(* IEC 61131-3 sources: TIA2AX/tests/V19/test_projects/expected/HW_2200330/ST80_PLC, 7 files *)

(* ---- HwIdentifiers.st ---- *)
TYPE
	HwIdentifiers : WORD
	(
		ST80_PLC_Profilschiene_0 :=	WORD#256,
		ST80_PLC :=	WORD#48,
		ST80_PLC_Card_reader_writer_1 :=	WORD#51,
		ST80_PLC_CPU_display_1 :=	WORD#54,
		ST80_PLC_OPC_UA_1 :=	WORD#117,
		ST80_PLC_DP_interface_1 :=	WORD#60,
		ST80_PLC_PROFINET_interface_1 :=	WORD#64,
		ST80_PLC_PROFINET_interface_1_Port_1 :=	WORD#65,
		ST80_PLC_PROFINET_interface_1_Port_2 :=	WORD#66,
		ST80_PLC_PROFINET_interface_2 :=	WORD#72,
		ST80_PLC_PROFINET_interface_2_Port_1 :=	WORD#73,
		ST80_Switch_SCALANCE_X_rack :=	WORD#412,
		ST80_Switch :=	WORD#413,
		ST80_Switch_ST80_Switch :=	WORD#414,
		ST80_Switch_SCALANCE_interface_1 :=	WORD#415,
		ST80_Switch_SCALANCE_interface_1_Port_1 :=	WORD#416,
		ST80_Switch_SCALANCE_interface_1_Port_2 :=	WORD#417,
		ST80_Switch_SCALANCE_interface_1_Port_3 :=	WORD#418,
		ST80_Switch_SCALANCE_interface_1_Port_4 :=	WORD#419,
		ST80_Switch_SCALANCE_interface_1_Port_5 :=	WORD#420,
		ST80_Switch_SCALANCE_interface_1_Port_6 :=	WORD#421,
		ST80_Switch_SCALANCE_interface_1_Port_7 :=	WORD#422,
		ST80_Switch_SCALANCE_interface_1_Port_8 :=	WORD#423,
		ST80_Switch_SCALANCE_interface_1_Port_9 :=	WORD#424,
		ST80_Switch_SCALANCE_interface_1_Port_10 :=	WORD#425,
		ST80_Switch_SCALANCE_interface_1_Port_11 :=	WORD#426,
		ST80_Switch_SCALANCE_interface_1_Port_12 :=	WORD#427,
		ST80_Switch_SCALANCE_interface_1_Port_13 :=	WORD#428,
		ST80_Switch_SCALANCE_interface_1_Port_14 :=	WORD#429,
		ST80_Switch_SCALANCE_interface_1_Port_15 :=	WORD#430,
		ST80_Switch_SCALANCE_interface_1_Port_16 :=	WORD#431,
		ST80_1_DM260_EB_Box_Rack :=	WORD#270,
		ST80_1_DM260_EB_Box :=	WORD#258,
		ST80_1_DM260_EB_Box_Interface :=	WORD#259,
		ST80_1_DM260_EB_Box_Interface_Port_1 :=	WORD#260,
		ST80_1_DM260_EB_Box_DataMan_260 :=	WORD#261,
		ST80_1_DM260_EB_Box_Acquisition_Control_1 :=	WORD#262,
		ST80_1_DM260_EB_Box_Acquisition_Status_1 :=	WORD#263,
		ST80_1_DM260_EB_Box_Results_Control_1 :=	WORD#264,
		ST80_1_DM260_EB_Box_Results_Status_1 :=	WORD#265,
		ST80_1_DM260_EB_Box_Soft_Event_Control_1 :=	WORD#266,
		ST80_1_DM260_EB_Box_User_Data_64_bytes_1 :=	WORD#267,
		ST80_1_DM260_EB_Box_Result_Data_64_bytes_1 :=	WORD#268,
		ST80_HMI_ConnectionBox_2_Connection_Box :=	WORD#272,
		ST80_HMI_ConnectionBox_2 :=	WORD#273,
		ST80_HMI_ConnectionBox_2_ST80_HMI_ConnectionBox_2 :=	WORD#274,
		ST80_HMI_ConnectionBox_2_SCALANCE_interface_1 :=	WORD#275,
		ST80_HMI_ConnectionBox_2_SCALANCE_interface_1_Port_1 :=	WORD#276,
		ST80_HMI_ConnectionBox_2_SCALANCE_interface_1_Port_2 :=	WORD#277,
		ST80_HMI_ConnectionBox_2_SCALANCE_interface_1_Port_3 :=	WORD#278,
		ST80_1_CMMT_1GF1_PN_IO_Interface :=	WORD#282,
		ST80_1_CMMT_1GF1_PN_IO_Interface_Port_1 :=	WORD#283,
		ST80_1_CMMT_1GF1_PN_IO_Interface_Port_2 :=	WORD#284,
		ST80_1_CMMT_1GF1_CMMT_AS_V1 :=	WORD#285,
		ST80_1_CMMT_1GF1_DO_SERVO_1_Module_Access_Point :=	WORD#287,
		ST80_1_CMMT_1GF1_DO_SERVO_1_Siemens_telegram_111_PZD_12_12 :=	WORD#288,
		ST80_1_CMMT_1GF1_Siemens_telegram_111_PZD_12_12 :=	WORD#288,
		ST80_1_CMMT_1GF2_PN_IO_Interface :=	WORD#292,
		ST80_1_CMMT_1GF2_PN_IO_Interface_Port_1 :=	WORD#293,
		ST80_1_CMMT_1GF2_PN_IO_Interface_Port_2 :=	WORD#294,
		ST80_1_CMMT_1GF2_CMMT_AS_V1 :=	WORD#295,
		ST80_1_CMMT_1GF2_DO_SERVO_1_Module_Access_Point :=	WORD#297,
		ST80_1_CMMT_1GF2_DO_SERVO_1_Siemens_telegram_111_PZD_12_12 :=	WORD#298,
		ST80_1_CMMT_1GF2_Siemens_telegram_111_PZD_12_12 :=	WORD#298,
		ST80_1_DM260_PB_Box_Rack :=	WORD#300,
		ST80_1_DM260_PB_Box :=	WORD#301,
		ST80_1_DM260_PB_Box_Interface :=	WORD#302,
		ST80_1_DM260_PB_Box_Interface_Port_1 :=	WORD#303,
		ST80_1_DM260_PB_Box_DataMan_260 :=	WORD#304,
		ST80_1_DM260_PB_Box_Acquisition_Control_1 :=	WORD#305,
		ST80_1_DM260_PB_Box_Acquisition_Status_1 :=	WORD#306,
		ST80_1_DM260_PB_Box_Results_Control_1 :=	WORD#307,
		ST80_1_DM260_PB_Box_Results_Status_1 :=	WORD#308,
		ST80_1_DM260_PB_Box_Soft_Event_Control_1 :=	WORD#309,
		ST80_1_DM260_PB_Box_User_Data_64_bytes_1 :=	WORD#310,
		ST80_1_DM260_PB_Box_Result_Data_64_bytes_1 :=	WORD#311,
		ST80_ET200SP_2_Rack_0 :=	WORD#313,
		ST80_ET200SP_2 :=	WORD#314,
		ST80_ET200SP_2_ST80_ET200SP_2 :=	WORD#315,
		ST80_ET200SP_2_PROFINET_interface :=	WORD#316,
		ST80_ET200SP_2_PROFINET_interface_Port_1 :=	WORD#318,
		ST80_ET200SP_2_PROFINET_interface_Port_2 :=	WORD#317,
		ST80_ET200SP_2_BA_2xRJ45 :=	WORD#318,
		ST80_ET200SP_2_BU_Cover_15_mm_1 :=	WORD#319,
		ST80_ET200SP_2_11M1 :=	WORD#320,
		ST80_ET200SP_2_11M2 :=	WORD#321,
		ST80_ET200SP_2_11M3 :=	WORD#322,
		ST80_ET200SP_2_11M4 :=	WORD#323,
		ST80_ET200SP_2_12M1 :=	WORD#324,
		ST80_ET200SP_2_12M2 :=	WORD#325,
		ST80_ET200SP_2_12M3 :=	WORD#326,
		ST80_ET200SP_2_12M4 :=	WORD#327,
		ST80_ET200SP_2_13M1 :=	WORD#328,
		ST80_ET200SP_2_13M2 :=	WORD#329,
		ST80_ET200SP_2_13M3 :=	WORD#330,
		ST80_ET200SP_2_13M4 :=	WORD#331,
		ST80_ET200SP_2_Servermodul_1 :=	WORD#332,
		ST80_1_TZ535_PN_Rack :=	WORD#334,
		ST80_1_TZ535_PN :=	WORD#335,
		ST80_1_TZ535_PN_Interface :=	WORD#336,
		ST80_1_TZ535_PN_Interface_Port_1 :=	WORD#337,
		ST80_1_TZ535_PN_Interface_Port_2 :=	WORD#338,
		ST80_1_TZ535_PN_2D_TZ535_PN_PROFINET_IO :=	WORD#339,
		ST80_1_TZ535_PN_In_Out_32_byte_1 :=	WORD#340,
		ST80_1_DM260_Housing_Rack :=	WORD#342,
		ST80_1_DM260_Housing :=	WORD#343,
		ST80_1_DM260_Housing_Interface :=	WORD#344,
		ST80_1_DM260_Housing_Interface_Port_1 :=	WORD#345,
		ST80_1_DM260_Housing_DataMan_260 :=	WORD#346,
		ST80_1_DM260_Housing_Acquisition_Control_1 :=	WORD#347,
		ST80_1_DM260_Housing_Acquisition_Status_1 :=	WORD#348,
		ST80_1_DM260_Housing_Results_Control_1 :=	WORD#349,
		ST80_1_DM260_Housing_Results_Status_1 :=	WORD#350,
		ST80_1_DM260_Housing_Soft_Event_Control_1 :=	WORD#351,
		ST80_1_DM260_Housing_User_Data_64_bytes_1 :=	WORD#352,
		ST80_1_DM260_Housing_Result_Data_64_bytes_1 :=	WORD#353,
		ST80_1_CMMT_3GF1_PN_IO_Interface :=	WORD#357,
		ST80_1_CMMT_3GF1_PN_IO_Interface_Port_1 :=	WORD#358,
		ST80_1_CMMT_3GF1_PN_IO_Interface_Port_2 :=	WORD#359,
		ST80_1_CMMT_3GF1_CMMT_AS_V1 :=	WORD#360,
		ST80_1_CMMT_3GF1_DO_SERVO_1_Module_Access_Point :=	WORD#362,
		ST80_1_CMMT_3GF1_DO_SERVO_1_Siemens_telegram_111_PZD_12_12 :=	WORD#363,
		ST80_1_CMMT_3GF1_Siemens_telegram_111_PZD_12_12 :=	WORD#363,
		ST80_CPX_PN_IO_Interface :=	WORD#367,
		ST80_CPX_PN_IO_Interface_Port_1 :=	WORD#368,
		ST80_CPX_PN_IO_Interface_Port_2 :=	WORD#369,
		ST80_CPX_CPX :=	WORD#370,
		ST80_CPX_MPA1S_VMPA1_FB_EMS_8_8DO_1 :=	WORD#371,
		ST80_CPX_MPA1S_VMPA1_FB_EMS_8_8DO_2 :=	WORD#372,
		ST80_CPX_MPA2S_VMPA2_FB_EMS_4_4DO_1 :=	WORD#373,
		ST80_CPX_MPA1S_VMPA1_FB_EMS_8_8DO_3 :=	WORD#374,
		ST80_CPX_MPA2S_VMPA2_FB_EMS_4_4DO_2 :=	WORD#375,
		ST80_CPX_MPA1S_VMPA1_FB_EMS_8_8DO_4 :=	WORD#376,
		ST80_CPX_MPA1S_VMPA1_FB_EMS_8_8DO_5 :=	WORD#377,
		ST80_CPX_MPA1G_VMPA1_FB_EMG_8_8DO_1 :=	WORD#378,
		ST80_CPX_MPA1G_VMPA1_FB_EMG_8_8DO_2 :=	WORD#379,
		ST80_CPX_MPA2G_VMPA2_FB_EMG_4_4DO_1 :=	WORD#380,
		ST80_CPX_MPA1G_VMPA1_FB_EMG_8_8DO_3 :=	WORD#381,
		ST80_CPX_MPA1G_VMPA1_FB_EMG_8_8DO_4 :=	WORD#382,
		ST80_CPX_MPA1G_VMPA1_FB_EMG_8_8DO_5 :=	WORD#383,
		ST80_CPX_MPA1G_VMPA1_FB_EMG_8_8DO_6 :=	WORD#384,
		ST80_ET200SP_Rack_0 :=	WORD#386,
		ST80_ET200SP :=	WORD#387,
		ST80_ET200SP_ST80_ET200SP :=	WORD#388,
		ST80_ET200SP_PROFINET_interface :=	WORD#389,
		ST80_ET200SP_PROFINET_interface_Port_1 :=	WORD#391,
		ST80_ET200SP_PROFINET_interface_Port_2 :=	WORD#390,
		ST80_ET200SP_BA_2xRJ45 :=	WORD#391,
		ST80_ET200SP_CM_4xIO_Link_1 :=	WORD#392,
		ST80_ET200SP_CM_4xIO_Link_2 :=	WORD#393,
		ST80_ET200SP_CM_4xIO_Link_3 :=	WORD#394,
		ST80_ET200SP_DI_16x24VDC_ST_1 :=	WORD#395,
		ST80_ET200SP_DI_16x24VDC_ST_2 :=	WORD#396,
		ST80_ET200SP_DI_16x24VDC_ST_3 :=	WORD#397,
		ST80_ET200SP_DI_16x24VDC_ST_4 :=	WORD#398,
		ST80_ET200SP_DQ_16x24VDC_0_5A_ST_1 :=	WORD#399,
		ST80_ET200SP_DQ_16x24VDC_0_5A_ST_2 :=	WORD#400,
		ST80_ET200SP_DQ_16x24VDC_0_5A_ST_3 :=	WORD#401,
		ST80_ET200SP_Servermodul_1 :=	WORD#402,
		ST80_HMI_ConnectionBox_Connection_Box :=	WORD#404,
		ST80_HMI_ConnectionBox :=	WORD#405,
		ST80_HMI_ConnectionBox_ST80_HMI_ConnectionBox :=	WORD#406,
		ST80_HMI_ConnectionBox_SCALANCE_interface_1 :=	WORD#407,
		ST80_HMI_ConnectionBox_SCALANCE_interface_1_Port_1 :=	WORD#408,
		ST80_HMI_ConnectionBox_SCALANCE_interface_1_Port_2 :=	WORD#409,
		ST80_HMI_ConnectionBox_SCALANCE_interface_1_Port_3 :=	WORD#410,
		NONE:= WORD#0
	);
END_TYPE

(* ---- HwInputs.st ---- *)
TYPE
	HwInputs : STRUCT
		ST80_1_DM260_EB_Box_Acquisition_Status_1 AT %B1205 : ARRAY[0..2] OF BYTE;
		ST80_1_DM260_EB_Box_Results_Status_1 AT %B1208 : BYTE;
		ST80_1_DM260_EB_Box_Soft_Event_Control_1 AT %B1209 : BYTE;
		ST80_1_DM260_EB_Box_Result_Data_64_bytes_1 AT %B1382 : ARRAY[0..71] OF BYTE;
		ST80_1_CMMT_1GF1_DO_SERVO_1_Siemens_telegram_111_PZD_12_12 AT %B1700 : ARRAY[0..23] OF BYTE;
		ST80_1_CMMT_1GF2_DO_SERVO_1_Siemens_telegram_111_PZD_12_12 AT %B1600 : ARRAY[0..23] OF BYTE;
		ST80_1_DM260_PB_Box_Acquisition_Status_1 AT %B1200 : ARRAY[0..2] OF BYTE;
		ST80_1_DM260_PB_Box_Results_Status_1 AT %B1203 : BYTE;
		ST80_1_DM260_PB_Box_Soft_Event_Control_1 AT %B1204 : BYTE;
		ST80_1_DM260_PB_Box_Result_Data_64_bytes_1 AT %B1210 : ARRAY[0..71] OF BYTE;
		ST80_ET200SP_2_11M1 AT %B600 : DWORD;
		ST80_ET200SP_2_11M2 AT %B604 : DWORD;
		ST80_ET200SP_2_11M3 AT %B608 : DWORD;
		ST80_ET200SP_2_11M4 AT %B612 : DWORD;
		ST80_ET200SP_2_12M1 AT %B616 : DWORD;
		ST80_ET200SP_2_12M2 AT %B620 : DWORD;
		ST80_ET200SP_2_12M3 AT %B624 : DWORD;
		ST80_ET200SP_2_12M4 AT %B628 : DWORD;
		ST80_ET200SP_2_13M1 AT %B632 : DWORD;
		ST80_ET200SP_2_13M2 AT %B636 : DWORD;
		ST80_ET200SP_2_13M3 AT %B640 : DWORD;
		ST80_ET200SP_2_13M4 AT %B644 : DWORD;
		ST80_1_TZ535_PN_In_Out_32_byte_1 AT %B1800 : ARRAY[0..31] OF BYTE;
		ST80_1_DM260_Housing_Acquisition_Status_1 AT %B1000 : ARRAY[0..2] OF BYTE;
		ST80_1_DM260_Housing_Results_Status_1 AT %B1003 : BYTE;
		ST80_1_DM260_Housing_Soft_Event_Control_1 AT %B1004 : BYTE;
		ST80_1_DM260_Housing_Result_Data_64_bytes_1 AT %B1010 : ARRAY[0..71] OF BYTE;
		ST80_1_CMMT_3GF1_DO_SERVO_1_Siemens_telegram_111_PZD_12_12 AT %B1500 : ARRAY[0..23] OF BYTE;
		ST80_ET200SP_CM_4xIO_Link_1 AT %B100 : ARRAY[0..31] OF BYTE;
		ST80_ET200SP_CM_4xIO_Link_2 AT %B132 : ARRAY[0..31] OF BYTE;
		ST80_ET200SP_CM_4xIO_Link_3 AT %B164 : ARRAY[0..31] OF BYTE;
		ST80_ET200SP_DI_16x24VDC_ST_1 AT %B0 : WORD;
		ST80_ET200SP_DI_16x24VDC_ST_2 AT %B2 : WORD;
		ST80_ET200SP_DI_16x24VDC_ST_3 AT %B4 : WORD;
		ST80_ET200SP_DI_16x24VDC_ST_4 AT %B6 : WORD;
	END_STRUCT;
END_TYPE

(* ---- HwOutputs.st ---- *)
TYPE
	HwOutputs : STRUCT
		ST80_1_DM260_EB_Box_Acquisition_Control_1 AT %B1201 : BYTE;
		ST80_1_DM260_EB_Box_Results_Control_1 AT %B1205 : BYTE;
		ST80_1_DM260_EB_Box_Soft_Event_Control_1 AT %B1206 : BYTE;
		ST80_1_DM260_EB_Box_User_Data_64_bytes_1 AT %B1378 : ARRAY[0..67] OF BYTE;
		ST80_1_CMMT_1GF1_DO_SERVO_1_Siemens_telegram_111_PZD_12_12 AT %B1700 : ARRAY[0..23] OF BYTE;
		ST80_1_CMMT_1GF2_DO_SERVO_1_Siemens_telegram_111_PZD_12_12 AT %B1600 : ARRAY[0..23] OF BYTE;
		ST80_1_DM260_PB_Box_Acquisition_Control_1 AT %B1200 : BYTE;
		ST80_1_DM260_PB_Box_Results_Control_1 AT %B1203 : BYTE;
		ST80_1_DM260_PB_Box_Soft_Event_Control_1 AT %B1204 : BYTE;
		ST80_1_DM260_PB_Box_User_Data_64_bytes_1 AT %B1210 : ARRAY[0..67] OF BYTE;
		ST80_ET200SP_2_11M1 AT %B600 : WORD;
		ST80_ET200SP_2_11M2 AT %B604 : WORD;
		ST80_ET200SP_2_11M3 AT %B608 : WORD;
		ST80_ET200SP_2_11M4 AT %B612 : WORD;
		ST80_ET200SP_2_12M1 AT %B616 : WORD;
		ST80_ET200SP_2_12M2 AT %B620 : WORD;
		ST80_ET200SP_2_12M3 AT %B624 : WORD;
		ST80_ET200SP_2_12M4 AT %B628 : WORD;
		ST80_ET200SP_2_13M1 AT %B632 : WORD;
		ST80_ET200SP_2_13M2 AT %B636 : WORD;
		ST80_ET200SP_2_13M3 AT %B640 : WORD;
		ST80_ET200SP_2_13M4 AT %B644 : WORD;
		ST80_1_TZ535_PN_In_Out_32_byte_1 AT %B1800 : ARRAY[0..31] OF BYTE;
		ST80_1_DM260_Housing_Acquisition_Control_1 AT %B1000 : BYTE;
		ST80_1_DM260_Housing_Results_Control_1 AT %B1003 : BYTE;
		ST80_1_DM260_Housing_Soft_Event_Control_1 AT %B1004 : BYTE;
		ST80_1_DM260_Housing_User_Data_64_bytes_1 AT %B1010 : ARRAY[0..67] OF BYTE;
		ST80_1_CMMT_3GF1_DO_SERVO_1_Siemens_telegram_111_PZD_12_12 AT %B1500 : ARRAY[0..23] OF BYTE;
		ST80_CPX_MPA1S_VMPA1_FB_EMS_8_8DO_1 AT %B200 : BYTE;
		ST80_CPX_MPA1S_VMPA1_FB_EMS_8_8DO_2 AT %B201 : BYTE;
		ST80_CPX_MPA2S_VMPA2_FB_EMS_4_4DO_1 AT %B202 : BYTE;
		ST80_CPX_MPA1S_VMPA1_FB_EMS_8_8DO_3 AT %B203 : BYTE;
		ST80_CPX_MPA2S_VMPA2_FB_EMS_4_4DO_2 AT %B204 : BYTE;
		ST80_CPX_MPA1S_VMPA1_FB_EMS_8_8DO_4 AT %B205 : BYTE;
		ST80_CPX_MPA1S_VMPA1_FB_EMS_8_8DO_5 AT %B206 : BYTE;
		ST80_CPX_MPA1G_VMPA1_FB_EMG_8_8DO_1 AT %B207 : BYTE;
		ST80_CPX_MPA1G_VMPA1_FB_EMG_8_8DO_2 AT %B208 : BYTE;
		ST80_CPX_MPA2G_VMPA2_FB_EMG_4_4DO_1 AT %B209 : BYTE;
		ST80_CPX_MPA1G_VMPA1_FB_EMG_8_8DO_3 AT %B210 : BYTE;
		ST80_CPX_MPA1G_VMPA1_FB_EMG_8_8DO_4 AT %B211 : BYTE;
		ST80_CPX_MPA1G_VMPA1_FB_EMG_8_8DO_5 AT %B212 : BYTE;
		ST80_CPX_MPA1G_VMPA1_FB_EMG_8_8DO_6 AT %B213 : BYTE;
		ST80_ET200SP_CM_4xIO_Link_1 AT %B100 : ARRAY[0..31] OF BYTE;
		ST80_ET200SP_CM_4xIO_Link_2 AT %B132 : ARRAY[0..31] OF BYTE;
		ST80_ET200SP_CM_4xIO_Link_3 AT %B164 : ARRAY[0..31] OF BYTE;
		ST80_ET200SP_DQ_16x24VDC_0_5A_ST_1 AT %B0 : WORD;
		ST80_ET200SP_DQ_16x24VDC_0_5A_ST_2 AT %B2 : WORD;
		ST80_ET200SP_DQ_16x24VDC_0_5A_ST_3 AT %B4 : WORD;
	END_STRUCT;
END_TYPE

(* ---- PlcInputs.st ---- *)
TYPE
	PlcInputs : STRUCT
		ST80_1_DM260_EB_Box_Acquisition_Status_1 : ARRAY[0..2] OF BYTE;
		ST80_1_DM260_EB_Box_Results_Status_1 : BYTE;
		ST80_1_DM260_EB_Box_Soft_Event_Control_1 : BYTE;
		ST80_1_DM260_EB_Box_Result_Data_64_bytes_1 : ARRAY[0..71] OF BYTE;
		ST80_1_CMMT_1GF1_DO_SERVO_1_Siemens_telegram_111_PZD_12_12 : ARRAY[0..23] OF BYTE;
		ST80_1_CMMT_1GF2_DO_SERVO_1_Siemens_telegram_111_PZD_12_12 : ARRAY[0..23] OF BYTE;
		ST80_1_DM260_PB_Box_Acquisition_Status_1 : ARRAY[0..2] OF BYTE;
		ST80_1_DM260_PB_Box_Results_Status_1 : BYTE;
		ST80_1_DM260_PB_Box_Soft_Event_Control_1 : BYTE;
		ST80_1_DM260_PB_Box_Result_Data_64_bytes_1 : ARRAY[0..71] OF BYTE;
		ST80_ET200SP_2_11M1 : DWORD;
		ST80_ET200SP_2_11M2 : DWORD;
		ST80_ET200SP_2_11M3 : DWORD;
		ST80_ET200SP_2_11M4 : DWORD;
		ST80_ET200SP_2_12M1 : DWORD;
		ST80_ET200SP_2_12M2 : DWORD;
		ST80_ET200SP_2_12M3 : DWORD;
		ST80_ET200SP_2_12M4 : DWORD;
		ST80_ET200SP_2_13M1 : DWORD;
		ST80_ET200SP_2_13M2 : DWORD;
		ST80_ET200SP_2_13M3 : DWORD;
		ST80_ET200SP_2_13M4 : DWORD;
		ST80_1_TZ535_PN_In_Out_32_byte_1 : ARRAY[0..31] OF BYTE;
		ST80_1_DM260_Housing_Acquisition_Status_1 : ARRAY[0..2] OF BYTE;
		ST80_1_DM260_Housing_Results_Status_1 : BYTE;
		ST80_1_DM260_Housing_Soft_Event_Control_1 : BYTE;
		ST80_1_DM260_Housing_Result_Data_64_bytes_1 : ARRAY[0..71] OF BYTE;
		ST80_1_CMMT_3GF1_DO_SERVO_1_Siemens_telegram_111_PZD_12_12 : ARRAY[0..23] OF BYTE;
		ST80_ET200SP_CM_4xIO_Link_1 : ARRAY[0..31] OF BYTE;
		ST80_ET200SP_CM_4xIO_Link_2 : ARRAY[0..31] OF BYTE;
		ST80_ET200SP_CM_4xIO_Link_3 : ARRAY[0..31] OF BYTE;
		ST80_ET200SP_DI_16x24VDC_ST_1 : WORD;
		ST80_ET200SP_DI_16x24VDC_ST_2 : WORD;
		ST80_ET200SP_DI_16x24VDC_ST_3 : WORD;
		ST80_ET200SP_DI_16x24VDC_ST_4 : WORD;
	END_STRUCT;
END_TYPE

(* ---- PlcOutputs.st ---- *)
TYPE
	PlcOutputs : STRUCT
		ST80_1_DM260_EB_Box_Acquisition_Control_1 : BYTE;
		ST80_1_DM260_EB_Box_Results_Control_1 : BYTE;
		ST80_1_DM260_EB_Box_Soft_Event_Control_1 : BYTE;
		ST80_1_DM260_EB_Box_User_Data_64_bytes_1 : ARRAY[0..67] OF BYTE;
		ST80_1_CMMT_1GF1_DO_SERVO_1_Siemens_telegram_111_PZD_12_12 : ARRAY[0..23] OF BYTE;
		ST80_1_CMMT_1GF2_DO_SERVO_1_Siemens_telegram_111_PZD_12_12 : ARRAY[0..23] OF BYTE;
		ST80_1_DM260_PB_Box_Acquisition_Control_1 : BYTE;
		ST80_1_DM260_PB_Box_Results_Control_1 : BYTE;
		ST80_1_DM260_PB_Box_Soft_Event_Control_1 : BYTE;
		ST80_1_DM260_PB_Box_User_Data_64_bytes_1 : ARRAY[0..67] OF BYTE;
		ST80_ET200SP_2_11M1 : WORD;
		ST80_ET200SP_2_11M2 : WORD;
		ST80_ET200SP_2_11M3 : WORD;
		ST80_ET200SP_2_11M4 : WORD;
		ST80_ET200SP_2_12M1 : WORD;
		ST80_ET200SP_2_12M2 : WORD;
		ST80_ET200SP_2_12M3 : WORD;
		ST80_ET200SP_2_12M4 : WORD;
		ST80_ET200SP_2_13M1 : WORD;
		ST80_ET200SP_2_13M2 : WORD;
		ST80_ET200SP_2_13M3 : WORD;
		ST80_ET200SP_2_13M4 : WORD;
		ST80_1_TZ535_PN_In_Out_32_byte_1 : ARRAY[0..31] OF BYTE;
		ST80_1_DM260_Housing_Acquisition_Control_1 : BYTE;
		ST80_1_DM260_Housing_Results_Control_1 : BYTE;
		ST80_1_DM260_Housing_Soft_Event_Control_1 : BYTE;
		ST80_1_DM260_Housing_User_Data_64_bytes_1 : ARRAY[0..67] OF BYTE;
		ST80_1_CMMT_3GF1_DO_SERVO_1_Siemens_telegram_111_PZD_12_12 : ARRAY[0..23] OF BYTE;
		ST80_CPX_MPA1S_VMPA1_FB_EMS_8_8DO_1 : BYTE;
		ST80_CPX_MPA1S_VMPA1_FB_EMS_8_8DO_2 : BYTE;
		ST80_CPX_MPA2S_VMPA2_FB_EMS_4_4DO_1 : BYTE;
		ST80_CPX_MPA1S_VMPA1_FB_EMS_8_8DO_3 : BYTE;
		ST80_CPX_MPA2S_VMPA2_FB_EMS_4_4DO_2 : BYTE;
		ST80_CPX_MPA1S_VMPA1_FB_EMS_8_8DO_4 : BYTE;
		ST80_CPX_MPA1S_VMPA1_FB_EMS_8_8DO_5 : BYTE;
		ST80_CPX_MPA1G_VMPA1_FB_EMG_8_8DO_1 : BYTE;
		ST80_CPX_MPA1G_VMPA1_FB_EMG_8_8DO_2 : BYTE;
		ST80_CPX_MPA2G_VMPA2_FB_EMG_4_4DO_1 : BYTE;
		ST80_CPX_MPA1G_VMPA1_FB_EMG_8_8DO_3 : BYTE;
		ST80_CPX_MPA1G_VMPA1_FB_EMG_8_8DO_4 : BYTE;
		ST80_CPX_MPA1G_VMPA1_FB_EMG_8_8DO_5 : BYTE;
		ST80_CPX_MPA1G_VMPA1_FB_EMG_8_8DO_6 : BYTE;
		ST80_ET200SP_CM_4xIO_Link_1 : ARRAY[0..31] OF BYTE;
		ST80_ET200SP_CM_4xIO_Link_2 : ARRAY[0..31] OF BYTE;
		ST80_ET200SP_CM_4xIO_Link_3 : ARRAY[0..31] OF BYTE;
		ST80_ET200SP_DQ_16x24VDC_0_5A_ST_1 : WORD;
		ST80_ET200SP_DQ_16x24VDC_0_5A_ST_2 : WORD;
		ST80_ET200SP_DQ_16x24VDC_0_5A_ST_3 : WORD;
	END_STRUCT;
END_TYPE

(* ---- CopyInputs.st ---- *)
FUNCTION CopyInputs
	VAR_EXTERNAL
		HwInputs : HwInputs;
		PlcInputs : PlcInputs;
	END_VAR
	PlcInputs.ST80_1_DM260_EB_Box_Acquisition_Status_1[0] := HwInputs.ST80_1_DM260_EB_Box_Acquisition_Status_1[0];
	PlcInputs.ST80_1_DM260_EB_Box_Acquisition_Status_1[1] := HwInputs.ST80_1_DM260_EB_Box_Acquisition_Status_1[1];
	PlcInputs.ST80_1_DM260_EB_Box_Acquisition_Status_1[2] := HwInputs.ST80_1_DM260_EB_Box_Acquisition_Status_1[2];
	PlcInputs.ST80_1_DM260_EB_Box_Results_Status_1 := HwInputs.ST80_1_DM260_EB_Box_Results_Status_1;
	PlcInputs.ST80_1_DM260_EB_Box_Soft_Event_Control_1 := HwInputs.ST80_1_DM260_EB_Box_Soft_Event_Control_1;
	PlcInputs.ST80_1_DM260_EB_Box_Result_Data_64_bytes_1[0] := HwInputs.ST80_1_DM260_EB_Box_Result_Data_64_bytes_1[0];
	PlcInputs.ST80_1_DM260_EB_Box_Result_Data_64_bytes_1[1] := HwInputs.ST80_1_DM260_EB_Box_Result_Data_64_bytes_1[1];
	PlcInputs.ST80_1_DM260_EB_Box_Result_Data_64_bytes_1[2] := HwInputs.ST80_1_DM260_EB_Box_Result_Data_64_bytes_1[2];
	PlcInputs.ST80_1_DM260_EB_Box_Result_Data_64_bytes_1[3] := HwInputs.ST80_1_DM260_EB_Box_Result_Data_64_bytes_1[3];
	PlcInputs.ST80_1_DM260_EB_Box_Result_Data_64_bytes_1[4] := HwInputs.ST80_1_DM260_EB_Box_Result_Data_64_bytes_1[4];
	PlcInputs.ST80_1_DM260_EB_Box_Result_Data_64_bytes_1[5] := HwInputs.ST80_1_DM260_EB_Box_Result_Data_64_bytes_1[5];
	PlcInputs.ST80_1_DM260_EB_Box_Result_Data_64_bytes_1[6] := HwInputs.ST80_1_DM260_EB_Box_Result_Data_64_bytes_1[6];
	PlcInputs.ST80_1_DM260_EB_Box_Result_Data_64_bytes_1[7] := HwInputs.ST80_1_DM260_EB_Box_Result_Data_64_bytes_1[7];
	PlcInputs.ST80_1_DM260_EB_Box_Result_Data_64_bytes_1[8] := HwInputs.ST80_1_DM260_EB_Box_Result_Data_64_bytes_1[8];
	PlcInputs.ST80_1_DM260_EB_Box_Result_Data_64_bytes_1[9] := HwInputs.ST80_1_DM260_EB_Box_Result_Data_64_bytes_1[9];
	PlcInputs.ST80_1_DM260_EB_Box_Result_Data_64_bytes_1[10] := HwInputs.ST80_1_DM260_EB_Box_Result_Data_64_bytes_1[10];
	PlcInputs.ST80_1_DM260_EB_Box_Result_Data_64_bytes_1[11] := HwInputs.ST80_1_DM260_EB_Box_Result_Data_64_bytes_1[11];
	PlcInputs.ST80_1_DM260_EB_Box_Result_Data_64_bytes_1[12] := HwInputs.ST80_1_DM260_EB_Box_Result_Data_64_bytes_1[12];
	PlcInputs.ST80_1_DM260_EB_Box_Result_Data_64_bytes_1[13] := HwInputs.ST80_1_DM260_EB_Box_Result_Data_64_bytes_1[13];
	PlcInputs.ST80_1_DM260_EB_Box_Result_Data_64_bytes_1[14] := HwInputs.ST80_1_DM260_EB_Box_Result_Data_64_bytes_1[14];
	PlcInputs.ST80_1_DM260_EB_Box_Result_Data_64_bytes_1[15] := HwInputs.ST80_1_DM260_EB_Box_Result_Data_64_bytes_1[15];
	PlcInputs.ST80_1_DM260_EB_Box_Result_Data_64_bytes_1[16] := HwInputs.ST80_1_DM260_EB_Box_Result_Data_64_bytes_1[16];
	PlcInputs.ST80_1_DM260_EB_Box_Result_Data_64_bytes_1[17] := HwInputs.ST80_1_DM260_EB_Box_Result_Data_64_bytes_1[17];
	PlcInputs.ST80_1_DM260_EB_Box_Result_Data_64_bytes_1[18] := HwInputs.ST80_1_DM260_EB_Box_Result_Data_64_bytes_1[18];
	PlcInputs.ST80_1_DM260_EB_Box_Result_Data_64_bytes_1[19] := HwInputs.ST80_1_DM260_EB_Box_Result_Data_64_bytes_1[19];
	PlcInputs.ST80_1_DM260_EB_Box_Result_Data_64_bytes_1[20] := HwInputs.ST80_1_DM260_EB_Box_Result_Data_64_bytes_1[20];
	PlcInputs.ST80_1_DM260_EB_Box_Result_Data_64_bytes_1[21] := HwInputs.ST80_1_DM260_EB_Box_Result_Data_64_bytes_1[21];
	PlcInputs.ST80_1_DM260_EB_Box_Result_Data_64_bytes_1[22] := HwInputs.ST80_1_DM260_EB_Box_Result_Data_64_bytes_1[22];
	PlcInputs.ST80_1_DM260_EB_Box_Result_Data_64_bytes_1[23] := HwInputs.ST80_1_DM260_EB_Box_Result_Data_64_bytes_1[23];
	PlcInputs.ST80_1_DM260_EB_Box_Result_Data_64_bytes_1[24] := HwInputs.ST80_1_DM260_EB_Box_Result_Data_64_bytes_1[24];
	PlcInputs.ST80_1_DM260_EB_Box_Result_Data_64_bytes_1[25] := HwInputs.ST80_1_DM260_EB_Box_Result_Data_64_bytes_1[25];
	PlcInputs.ST80_1_DM260_EB_Box_Result_Data_64_bytes_1[26] := HwInputs.ST80_1_DM260_EB_Box_Result_Data_64_bytes_1[26];
	PlcInputs.ST80_1_DM260_EB_Box_Result_Data_64_bytes_1[27] := HwInputs.ST80_1_DM260_EB_Box_Result_Data_64_bytes_1[27];
	PlcInputs.ST80_1_DM260_EB_Box_Result_Data_64_bytes_1[28] := HwInputs.ST80_1_DM260_EB_Box_Result_Data_64_bytes_1[28];
	PlcInputs.ST80_1_DM260_EB_Box_Result_Data_64_bytes_1[29] := HwInputs.ST80_1_DM260_EB_Box_Result_Data_64_bytes_1[29];
	PlcInputs.ST80_1_DM260_EB_Box_Result_Data_64_bytes_1[30] := HwInputs.ST80_1_DM260_EB_Box_Result_Data_64_bytes_1[30];
	PlcInputs.ST80_1_DM260_EB_Box_Result_Data_64_bytes_1[31] := HwInputs.ST80_1_DM260_EB_Box_Result_Data_64_bytes_1[31];
	PlcInputs.ST80_1_DM260_EB_Box_Result_Data_64_bytes_1[32] := HwInputs.ST80_1_DM260_EB_Box_Result_Data_64_bytes_1[32];
	PlcInputs.ST80_1_DM260_EB_Box_Result_Data_64_bytes_1[33] := HwInputs.ST80_1_DM260_EB_Box_Result_Data_64_bytes_1[33];
	PlcInputs.ST80_1_DM260_EB_Box_Result_Data_64_bytes_1[34] := HwInputs.ST80_1_DM260_EB_Box_Result_Data_64_bytes_1[34];
	PlcInputs.ST80_1_DM260_EB_Box_Result_Data_64_bytes_1[35] := HwInputs.ST80_1_DM260_EB_Box_Result_Data_64_bytes_1[35];
	PlcInputs.ST80_1_DM260_EB_Box_Result_Data_64_bytes_1[36] := HwInputs.ST80_1_DM260_EB_Box_Result_Data_64_bytes_1[36];
	PlcInputs.ST80_1_DM260_EB_Box_Result_Data_64_bytes_1[37] := HwInputs.ST80_1_DM260_EB_Box_Result_Data_64_bytes_1[37];
	PlcInputs.ST80_1_DM260_EB_Box_Result_Data_64_bytes_1[38] := HwInputs.ST80_1_DM260_EB_Box_Result_Data_64_bytes_1[38];
	PlcInputs.ST80_1_DM260_EB_Box_Result_Data_64_bytes_1[39] := HwInputs.ST80_1_DM260_EB_Box_Result_Data_64_bytes_1[39];
	PlcInputs.ST80_1_DM260_EB_Box_Result_Data_64_bytes_1[40] := HwInputs.ST80_1_DM260_EB_Box_Result_Data_64_bytes_1[40];
	PlcInputs.ST80_1_DM260_EB_Box_Result_Data_64_bytes_1[41] := HwInputs.ST80_1_DM260_EB_Box_Result_Data_64_bytes_1[41];
	PlcInputs.ST80_1_DM260_EB_Box_Result_Data_64_bytes_1[42] := HwInputs.ST80_1_DM260_EB_Box_Result_Data_64_bytes_1[42];
	PlcInputs.ST80_1_DM260_EB_Box_Result_Data_64_bytes_1[43] := HwInputs.ST80_1_DM260_EB_Box_Result_Data_64_bytes_1[43];
	PlcInputs.ST80_1_DM260_EB_Box_Result_Data_64_bytes_1[44] := HwInputs.ST80_1_DM260_EB_Box_Result_Data_64_bytes_1[44];
	PlcInputs.ST80_1_DM260_EB_Box_Result_Data_64_bytes_1[45] := HwInputs.ST80_1_DM260_EB_Box_Result_Data_64_bytes_1[45];
	PlcInputs.ST80_1_DM260_EB_Box_Result_Data_64_bytes_1[46] := HwInputs.ST80_1_DM260_EB_Box_Result_Data_64_bytes_1[46];
	PlcInputs.ST80_1_DM260_EB_Box_Result_Data_64_bytes_1[47] := HwInputs.ST80_1_DM260_EB_Box_Result_Data_64_bytes_1[47];
	PlcInputs.ST80_1_DM260_EB_Box_Result_Data_64_bytes_1[48] := HwInputs.ST80_1_DM260_EB_Box_Result_Data_64_bytes_1[48];
	PlcInputs.ST80_1_DM260_EB_Box_Result_Data_64_bytes_1[49] := HwInputs.ST80_1_DM260_EB_Box_Result_Data_64_bytes_1[49];
	PlcInputs.ST80_1_DM260_EB_Box_Result_Data_64_bytes_1[50] := HwInputs.ST80_1_DM260_EB_Box_Result_Data_64_bytes_1[50];
	PlcInputs.ST80_1_DM260_EB_Box_Result_Data_64_bytes_1[51] := HwInputs.ST80_1_DM260_EB_Box_Result_Data_64_bytes_1[51];
	PlcInputs.ST80_1_DM260_EB_Box_Result_Data_64_bytes_1[52] := HwInputs.ST80_1_DM260_EB_Box_Result_Data_64_bytes_1[52];
	PlcInputs.ST80_1_DM260_EB_Box_Result_Data_64_bytes_1[53] := HwInputs.ST80_1_DM260_EB_Box_Result_Data_64_bytes_1[53];
	PlcInputs.ST80_1_DM260_EB_Box_Result_Data_64_bytes_1[54] := HwInputs.ST80_1_DM260_EB_Box_Result_Data_64_bytes_1[54];
	PlcInputs.ST80_1_DM260_EB_Box_Result_Data_64_bytes_1[55] := HwInputs.ST80_1_DM260_EB_Box_Result_Data_64_bytes_1[55];
	PlcInputs.ST80_1_DM260_EB_Box_Result_Data_64_bytes_1[56] := HwInputs.ST80_1_DM260_EB_Box_Result_Data_64_bytes_1[56];
	PlcInputs.ST80_1_DM260_EB_Box_Result_Data_64_bytes_1[57] := HwInputs.ST80_1_DM260_EB_Box_Result_Data_64_bytes_1[57];
	PlcInputs.ST80_1_DM260_EB_Box_Result_Data_64_bytes_1[58] := HwInputs.ST80_1_DM260_EB_Box_Result_Data_64_bytes_1[58];
	PlcInputs.ST80_1_DM260_EB_Box_Result_Data_64_bytes_1[59] := HwInputs.ST80_1_DM260_EB_Box_Result_Data_64_bytes_1[59];
	PlcInputs.ST80_1_DM260_EB_Box_Result_Data_64_bytes_1[60] := HwInputs.ST80_1_DM260_EB_Box_Result_Data_64_bytes_1[60];
	PlcInputs.ST80_1_DM260_EB_Box_Result_Data_64_bytes_1[61] := HwInputs.ST80_1_DM260_EB_Box_Result_Data_64_bytes_1[61];
	PlcInputs.ST80_1_DM260_EB_Box_Result_Data_64_bytes_1[62] := HwInputs.ST80_1_DM260_EB_Box_Result_Data_64_bytes_1[62];
	PlcInputs.ST80_1_DM260_EB_Box_Result_Data_64_bytes_1[63] := HwInputs.ST80_1_DM260_EB_Box_Result_Data_64_bytes_1[63];
	PlcInputs.ST80_1_DM260_EB_Box_Result_Data_64_bytes_1[64] := HwInputs.ST80_1_DM260_EB_Box_Result_Data_64_bytes_1[64];
	PlcInputs.ST80_1_DM260_EB_Box_Result_Data_64_bytes_1[65] := HwInputs.ST80_1_DM260_EB_Box_Result_Data_64_bytes_1[65];
	PlcInputs.ST80_1_DM260_EB_Box_Result_Data_64_bytes_1[66] := HwInputs.ST80_1_DM260_EB_Box_Result_Data_64_bytes_1[66];
	PlcInputs.ST80_1_DM260_EB_Box_Result_Data_64_bytes_1[67] := HwInputs.ST80_1_DM260_EB_Box_Result_Data_64_bytes_1[67];
	PlcInputs.ST80_1_DM260_EB_Box_Result_Data_64_bytes_1[68] := HwInputs.ST80_1_DM260_EB_Box_Result_Data_64_bytes_1[68];
	PlcInputs.ST80_1_DM260_EB_Box_Result_Data_64_bytes_1[69] := HwInputs.ST80_1_DM260_EB_Box_Result_Data_64_bytes_1[69];
	PlcInputs.ST80_1_DM260_EB_Box_Result_Data_64_bytes_1[70] := HwInputs.ST80_1_DM260_EB_Box_Result_Data_64_bytes_1[70];
	PlcInputs.ST80_1_DM260_EB_Box_Result_Data_64_bytes_1[71] := HwInputs.ST80_1_DM260_EB_Box_Result_Data_64_bytes_1[71];
	PlcInputs.ST80_1_CMMT_1GF1_DO_SERVO_1_Siemens_telegram_111_PZD_12_12[0] := HwInputs.ST80_1_CMMT_1GF1_DO_SERVO_1_Siemens_telegram_111_PZD_12_12[0];
	PlcInputs.ST80_1_CMMT_1GF1_DO_SERVO_1_Siemens_telegram_111_PZD_12_12[1] := HwInputs.ST80_1_CMMT_1GF1_DO_SERVO_1_Siemens_telegram_111_PZD_12_12[1];
	PlcInputs.ST80_1_CMMT_1GF1_DO_SERVO_1_Siemens_telegram_111_PZD_12_12[2] := HwInputs.ST80_1_CMMT_1GF1_DO_SERVO_1_Siemens_telegram_111_PZD_12_12[2];
	PlcInputs.ST80_1_CMMT_1GF1_DO_SERVO_1_Siemens_telegram_111_PZD_12_12[3] := HwInputs.ST80_1_CMMT_1GF1_DO_SERVO_1_Siemens_telegram_111_PZD_12_12[3];
	PlcInputs.ST80_1_CMMT_1GF1_DO_SERVO_1_Siemens_telegram_111_PZD_12_12[4] := HwInputs.ST80_1_CMMT_1GF1_DO_SERVO_1_Siemens_telegram_111_PZD_12_12[4];
	PlcInputs.ST80_1_CMMT_1GF1_DO_SERVO_1_Siemens_telegram_111_PZD_12_12[5] := HwInputs.ST80_1_CMMT_1GF1_DO_SERVO_1_Siemens_telegram_111_PZD_12_12[5];
	PlcInputs.ST80_1_CMMT_1GF1_DO_SERVO_1_Siemens_telegram_111_PZD_12_12[6] := HwInputs.ST80_1_CMMT_1GF1_DO_SERVO_1_Siemens_telegram_111_PZD_12_12[6];
	PlcInputs.ST80_1_CMMT_1GF1_DO_SERVO_1_Siemens_telegram_111_PZD_12_12[7] := HwInputs.ST80_1_CMMT_1GF1_DO_SERVO_1_Siemens_telegram_111_PZD_12_12[7];
	PlcInputs.ST80_1_CMMT_1GF1_DO_SERVO_1_Siemens_telegram_111_PZD_12_12[8] := HwInputs.ST80_1_CMMT_1GF1_DO_SERVO_1_Siemens_telegram_111_PZD_12_12[8];
	PlcInputs.ST80_1_CMMT_1GF1_DO_SERVO_1_Siemens_telegram_111_PZD_12_12[9] := HwInputs.ST80_1_CMMT_1GF1_DO_SERVO_1_Siemens_telegram_111_PZD_12_12[9];
	PlcInputs.ST80_1_CMMT_1GF1_DO_SERVO_1_Siemens_telegram_111_PZD_12_12[10] := HwInputs.ST80_1_CMMT_1GF1_DO_SERVO_1_Siemens_telegram_111_PZD_12_12[10];
	PlcInputs.ST80_1_CMMT_1GF1_DO_SERVO_1_Siemens_telegram_111_PZD_12_12[11] := HwInputs.ST80_1_CMMT_1GF1_DO_SERVO_1_Siemens_telegram_111_PZD_12_12[11];
	PlcInputs.ST80_1_CMMT_1GF1_DO_SERVO_1_Siemens_telegram_111_PZD_12_12[12] := HwInputs.ST80_1_CMMT_1GF1_DO_SERVO_1_Siemens_telegram_111_PZD_12_12[12];
	PlcInputs.ST80_1_CMMT_1GF1_DO_SERVO_1_Siemens_telegram_111_PZD_12_12[13] := HwInputs.ST80_1_CMMT_1GF1_DO_SERVO_1_Siemens_telegram_111_PZD_12_12[13];
	PlcInputs.ST80_1_CMMT_1GF1_DO_SERVO_1_Siemens_telegram_111_PZD_12_12[14] := HwInputs.ST80_1_CMMT_1GF1_DO_SERVO_1_Siemens_telegram_111_PZD_12_12[14];
	PlcInputs.ST80_1_CMMT_1GF1_DO_SERVO_1_Siemens_telegram_111_PZD_12_12[15] := HwInputs.ST80_1_CMMT_1GF1_DO_SERVO_1_Siemens_telegram_111_PZD_12_12[15];
	PlcInputs.ST80_1_CMMT_1GF1_DO_SERVO_1_Siemens_telegram_111_PZD_12_12[16] := HwInputs.ST80_1_CMMT_1GF1_DO_SERVO_1_Siemens_telegram_111_PZD_12_12[16];
	PlcInputs.ST80_1_CMMT_1GF1_DO_SERVO_1_Siemens_telegram_111_PZD_12_12[17] := HwInputs.ST80_1_CMMT_1GF1_DO_SERVO_1_Siemens_telegram_111_PZD_12_12[17];
	PlcInputs.ST80_1_CMMT_1GF1_DO_SERVO_1_Siemens_telegram_111_PZD_12_12[18] := HwInputs.ST80_1_CMMT_1GF1_DO_SERVO_1_Siemens_telegram_111_PZD_12_12[18];
	PlcInputs.ST80_1_CMMT_1GF1_DO_SERVO_1_Siemens_telegram_111_PZD_12_12[19] := HwInputs.ST80_1_CMMT_1GF1_DO_SERVO_1_Siemens_telegram_111_PZD_12_12[19];
	PlcInputs.ST80_1_CMMT_1GF1_DO_SERVO_1_Siemens_telegram_111_PZD_12_12[20] := HwInputs.ST80_1_CMMT_1GF1_DO_SERVO_1_Siemens_telegram_111_PZD_12_12[20];
	PlcInputs.ST80_1_CMMT_1GF1_DO_SERVO_1_Siemens_telegram_111_PZD_12_12[21] := HwInputs.ST80_1_CMMT_1GF1_DO_SERVO_1_Siemens_telegram_111_PZD_12_12[21];
	PlcInputs.ST80_1_CMMT_1GF1_DO_SERVO_1_Siemens_telegram_111_PZD_12_12[22] := HwInputs.ST80_1_CMMT_1GF1_DO_SERVO_1_Siemens_telegram_111_PZD_12_12[22];
	PlcInputs.ST80_1_CMMT_1GF1_DO_SERVO_1_Siemens_telegram_111_PZD_12_12[23] := HwInputs.ST80_1_CMMT_1GF1_DO_SERVO_1_Siemens_telegram_111_PZD_12_12[23];
	PlcInputs.ST80_1_CMMT_1GF2_DO_SERVO_1_Siemens_telegram_111_PZD_12_12[0] := HwInputs.ST80_1_CMMT_1GF2_DO_SERVO_1_Siemens_telegram_111_PZD_12_12[0];
	PlcInputs.ST80_1_CMMT_1GF2_DO_SERVO_1_Siemens_telegram_111_PZD_12_12[1] := HwInputs.ST80_1_CMMT_1GF2_DO_SERVO_1_Siemens_telegram_111_PZD_12_12[1];
	PlcInputs.ST80_1_CMMT_1GF2_DO_SERVO_1_Siemens_telegram_111_PZD_12_12[2] := HwInputs.ST80_1_CMMT_1GF2_DO_SERVO_1_Siemens_telegram_111_PZD_12_12[2];
	PlcInputs.ST80_1_CMMT_1GF2_DO_SERVO_1_Siemens_telegram_111_PZD_12_12[3] := HwInputs.ST80_1_CMMT_1GF2_DO_SERVO_1_Siemens_telegram_111_PZD_12_12[3];
	PlcInputs.ST80_1_CMMT_1GF2_DO_SERVO_1_Siemens_telegram_111_PZD_12_12[4] := HwInputs.ST80_1_CMMT_1GF2_DO_SERVO_1_Siemens_telegram_111_PZD_12_12[4];
	PlcInputs.ST80_1_CMMT_1GF2_DO_SERVO_1_Siemens_telegram_111_PZD_12_12[5] := HwInputs.ST80_1_CMMT_1GF2_DO_SERVO_1_Siemens_telegram_111_PZD_12_12[5];
	PlcInputs.ST80_1_CMMT_1GF2_DO_SERVO_1_Siemens_telegram_111_PZD_12_12[6] := HwInputs.ST80_1_CMMT_1GF2_DO_SERVO_1_Siemens_telegram_111_PZD_12_12[6];
	PlcInputs.ST80_1_CMMT_1GF2_DO_SERVO_1_Siemens_telegram_111_PZD_12_12[7] := HwInputs.ST80_1_CMMT_1GF2_DO_SERVO_1_Siemens_telegram_111_PZD_12_12[7];
	PlcInputs.ST80_1_CMMT_1GF2_DO_SERVO_1_Siemens_telegram_111_PZD_12_12[8] := HwInputs.ST80_1_CMMT_1GF2_DO_SERVO_1_Siemens_telegram_111_PZD_12_12[8];
	PlcInputs.ST80_1_CMMT_1GF2_DO_SERVO_1_Siemens_telegram_111_PZD_12_12[9] := HwInputs.ST80_1_CMMT_1GF2_DO_SERVO_1_Siemens_telegram_111_PZD_12_12[9];
	PlcInputs.ST80_1_CMMT_1GF2_DO_SERVO_1_Siemens_telegram_111_PZD_12_12[10] := HwInputs.ST80_1_CMMT_1GF2_DO_SERVO_1_Siemens_telegram_111_PZD_12_12[10];
	PlcInputs.ST80_1_CMMT_1GF2_DO_SERVO_1_Siemens_telegram_111_PZD_12_12[11] := HwInputs.ST80_1_CMMT_1GF2_DO_SERVO_1_Siemens_telegram_111_PZD_12_12[11];
	PlcInputs.ST80_1_CMMT_1GF2_DO_SERVO_1_Siemens_telegram_111_PZD_12_12[12] := HwInputs.ST80_1_CMMT_1GF2_DO_SERVO_1_Siemens_telegram_111_PZD_12_12[12];
	PlcInputs.ST80_1_CMMT_1GF2_DO_SERVO_1_Siemens_telegram_111_PZD_12_12[13] := HwInputs.ST80_1_CMMT_1GF2_DO_SERVO_1_Siemens_telegram_111_PZD_12_12[13];
	PlcInputs.ST80_1_CMMT_1GF2_DO_SERVO_1_Siemens_telegram_111_PZD_12_12[14] := HwInputs.ST80_1_CMMT_1GF2_DO_SERVO_1_Siemens_telegram_111_PZD_12_12[14];
	PlcInputs.ST80_1_CMMT_1GF2_DO_SERVO_1_Siemens_telegram_111_PZD_12_12[15] := HwInputs.ST80_1_CMMT_1GF2_DO_SERVO_1_Siemens_telegram_111_PZD_12_12[15];
	PlcInputs.ST80_1_CMMT_1GF2_DO_SERVO_1_Siemens_telegram_111_PZD_12_12[16] := HwInputs.ST80_1_CMMT_1GF2_DO_SERVO_1_Siemens_telegram_111_PZD_12_12[16];
	PlcInputs.ST80_1_CMMT_1GF2_DO_SERVO_1_Siemens_telegram_111_PZD_12_12[17] := HwInputs.ST80_1_CMMT_1GF2_DO_SERVO_1_Siemens_telegram_111_PZD_12_12[17];
	PlcInputs.ST80_1_CMMT_1GF2_DO_SERVO_1_Siemens_telegram_111_PZD_12_12[18] := HwInputs.ST80_1_CMMT_1GF2_DO_SERVO_1_Siemens_telegram_111_PZD_12_12[18];
	PlcInputs.ST80_1_CMMT_1GF2_DO_SERVO_1_Siemens_telegram_111_PZD_12_12[19] := HwInputs.ST80_1_CMMT_1GF2_DO_SERVO_1_Siemens_telegram_111_PZD_12_12[19];
	PlcInputs.ST80_1_CMMT_1GF2_DO_SERVO_1_Siemens_telegram_111_PZD_12_12[20] := HwInputs.ST80_1_CMMT_1GF2_DO_SERVO_1_Siemens_telegram_111_PZD_12_12[20];
	PlcInputs.ST80_1_CMMT_1GF2_DO_SERVO_1_Siemens_telegram_111_PZD_12_12[21] := HwInputs.ST80_1_CMMT_1GF2_DO_SERVO_1_Siemens_telegram_111_PZD_12_12[21];
	PlcInputs.ST80_1_CMMT_1GF2_DO_SERVO_1_Siemens_telegram_111_PZD_12_12[22] := HwInputs.ST80_1_CMMT_1GF2_DO_SERVO_1_Siemens_telegram_111_PZD_12_12[22];
	PlcInputs.ST80_1_CMMT_1GF2_DO_SERVO_1_Siemens_telegram_111_PZD_12_12[23] := HwInputs.ST80_1_CMMT_1GF2_DO_SERVO_1_Siemens_telegram_111_PZD_12_12[23];
	PlcInputs.ST80_1_DM260_PB_Box_Acquisition_Status_1[0] := HwInputs.ST80_1_DM260_PB_Box_Acquisition_Status_1[0];
	PlcInputs.ST80_1_DM260_PB_Box_Acquisition_Status_1[1] := HwInputs.ST80_1_DM260_PB_Box_Acquisition_Status_1[1];
	PlcInputs.ST80_1_DM260_PB_Box_Acquisition_Status_1[2] := HwInputs.ST80_1_DM260_PB_Box_Acquisition_Status_1[2];
	PlcInputs.ST80_1_DM260_PB_Box_Results_Status_1 := HwInputs.ST80_1_DM260_PB_Box_Results_Status_1;
	PlcInputs.ST80_1_DM260_PB_Box_Soft_Event_Control_1 := HwInputs.ST80_1_DM260_PB_Box_Soft_Event_Control_1;
	PlcInputs.ST80_1_DM260_PB_Box_Result_Data_64_bytes_1[0] := HwInputs.ST80_1_DM260_PB_Box_Result_Data_64_bytes_1[0];
	PlcInputs.ST80_1_DM260_PB_Box_Result_Data_64_bytes_1[1] := HwInputs.ST80_1_DM260_PB_Box_Result_Data_64_bytes_1[1];
	PlcInputs.ST80_1_DM260_PB_Box_Result_Data_64_bytes_1[2] := HwInputs.ST80_1_DM260_PB_Box_Result_Data_64_bytes_1[2];
	PlcInputs.ST80_1_DM260_PB_Box_Result_Data_64_bytes_1[3] := HwInputs.ST80_1_DM260_PB_Box_Result_Data_64_bytes_1[3];
	PlcInputs.ST80_1_DM260_PB_Box_Result_Data_64_bytes_1[4] := HwInputs.ST80_1_DM260_PB_Box_Result_Data_64_bytes_1[4];
	PlcInputs.ST80_1_DM260_PB_Box_Result_Data_64_bytes_1[5] := HwInputs.ST80_1_DM260_PB_Box_Result_Data_64_bytes_1[5];
	PlcInputs.ST80_1_DM260_PB_Box_Result_Data_64_bytes_1[6] := HwInputs.ST80_1_DM260_PB_Box_Result_Data_64_bytes_1[6];
	PlcInputs.ST80_1_DM260_PB_Box_Result_Data_64_bytes_1[7] := HwInputs.ST80_1_DM260_PB_Box_Result_Data_64_bytes_1[7];
	PlcInputs.ST80_1_DM260_PB_Box_Result_Data_64_bytes_1[8] := HwInputs.ST80_1_DM260_PB_Box_Result_Data_64_bytes_1[8];
	PlcInputs.ST80_1_DM260_PB_Box_Result_Data_64_bytes_1[9] := HwInputs.ST80_1_DM260_PB_Box_Result_Data_64_bytes_1[9];
	PlcInputs.ST80_1_DM260_PB_Box_Result_Data_64_bytes_1[10] := HwInputs.ST80_1_DM260_PB_Box_Result_Data_64_bytes_1[10];
	PlcInputs.ST80_1_DM260_PB_Box_Result_Data_64_bytes_1[11] := HwInputs.ST80_1_DM260_PB_Box_Result_Data_64_bytes_1[11];
	PlcInputs.ST80_1_DM260_PB_Box_Result_Data_64_bytes_1[12] := HwInputs.ST80_1_DM260_PB_Box_Result_Data_64_bytes_1[12];
	PlcInputs.ST80_1_DM260_PB_Box_Result_Data_64_bytes_1[13] := HwInputs.ST80_1_DM260_PB_Box_Result_Data_64_bytes_1[13];
	PlcInputs.ST80_1_DM260_PB_Box_Result_Data_64_bytes_1[14] := HwInputs.ST80_1_DM260_PB_Box_Result_Data_64_bytes_1[14];
	PlcInputs.ST80_1_DM260_PB_Box_Result_Data_64_bytes_1[15] := HwInputs.ST80_1_DM260_PB_Box_Result_Data_64_bytes_1[15];
	PlcInputs.ST80_1_DM260_PB_Box_Result_Data_64_bytes_1[16] := HwInputs.ST80_1_DM260_PB_Box_Result_Data_64_bytes_1[16];
	PlcInputs.ST80_1_DM260_PB_Box_Result_Data_64_bytes_1[17] := HwInputs.ST80_1_DM260_PB_Box_Result_Data_64_bytes_1[17];
	PlcInputs.ST80_1_DM260_PB_Box_Result_Data_64_bytes_1[18] := HwInputs.ST80_1_DM260_PB_Box_Result_Data_64_bytes_1[18];
	PlcInputs.ST80_1_DM260_PB_Box_Result_Data_64_bytes_1[19] := HwInputs.ST80_1_DM260_PB_Box_Result_Data_64_bytes_1[19];
	PlcInputs.ST80_1_DM260_PB_Box_Result_Data_64_bytes_1[20] := HwInputs.ST80_1_DM260_PB_Box_Result_Data_64_bytes_1[20];
	PlcInputs.ST80_1_DM260_PB_Box_Result_Data_64_bytes_1[21] := HwInputs.ST80_1_DM260_PB_Box_Result_Data_64_bytes_1[21];
	PlcInputs.ST80_1_DM260_PB_Box_Result_Data_64_bytes_1[22] := HwInputs.ST80_1_DM260_PB_Box_Result_Data_64_bytes_1[22];
	PlcInputs.ST80_1_DM260_PB_Box_Result_Data_64_bytes_1[23] := HwInputs.ST80_1_DM260_PB_Box_Result_Data_64_bytes_1[23];
	PlcInputs.ST80_1_DM260_PB_Box_Result_Data_64_bytes_1[24] := HwInputs.ST80_1_DM260_PB_Box_Result_Data_64_bytes_1[24];
	PlcInputs.ST80_1_DM260_PB_Box_Result_Data_64_bytes_1[25] := HwInputs.ST80_1_DM260_PB_Box_Result_Data_64_bytes_1[25];
	PlcInputs.ST80_1_DM260_PB_Box_Result_Data_64_bytes_1[26] := HwInputs.ST80_1_DM260_PB_Box_Result_Data_64_bytes_1[26];
	PlcInputs.ST80_1_DM260_PB_Box_Result_Data_64_bytes_1[27] := HwInputs.ST80_1_DM260_PB_Box_Result_Data_64_bytes_1[27];
	PlcInputs.ST80_1_DM260_PB_Box_Result_Data_64_bytes_1[28] := HwInputs.ST80_1_DM260_PB_Box_Result_Data_64_bytes_1[28];
	PlcInputs.ST80_1_DM260_PB_Box_Result_Data_64_bytes_1[29] := HwInputs.ST80_1_DM260_PB_Box_Result_Data_64_bytes_1[29];
	PlcInputs.ST80_1_DM260_PB_Box_Result_Data_64_bytes_1[30] := HwInputs.ST80_1_DM260_PB_Box_Result_Data_64_bytes_1[30];
	PlcInputs.ST80_1_DM260_PB_Box_Result_Data_64_bytes_1[31] := HwInputs.ST80_1_DM260_PB_Box_Result_Data_64_bytes_1[31];
	PlcInputs.ST80_1_DM260_PB_Box_Result_Data_64_bytes_1[32] := HwInputs.ST80_1_DM260_PB_Box_Result_Data_64_bytes_1[32];
	PlcInputs.ST80_1_DM260_PB_Box_Result_Data_64_bytes_1[33] := HwInputs.ST80_1_DM260_PB_Box_Result_Data_64_bytes_1[33];
	PlcInputs.ST80_1_DM260_PB_Box_Result_Data_64_bytes_1[34] := HwInputs.ST80_1_DM260_PB_Box_Result_Data_64_bytes_1[34];
	PlcInputs.ST80_1_DM260_PB_Box_Result_Data_64_bytes_1[35] := HwInputs.ST80_1_DM260_PB_Box_Result_Data_64_bytes_1[35];
	PlcInputs.ST80_1_DM260_PB_Box_Result_Data_64_bytes_1[36] := HwInputs.ST80_1_DM260_PB_Box_Result_Data_64_bytes_1[36];
	PlcInputs.ST80_1_DM260_PB_Box_Result_Data_64_bytes_1[37] := HwInputs.ST80_1_DM260_PB_Box_Result_Data_64_bytes_1[37];
	PlcInputs.ST80_1_DM260_PB_Box_Result_Data_64_bytes_1[38] := HwInputs.ST80_1_DM260_PB_Box_Result_Data_64_bytes_1[38];
	PlcInputs.ST80_1_DM260_PB_Box_Result_Data_64_bytes_1[39] := HwInputs.ST80_1_DM260_PB_Box_Result_Data_64_bytes_1[39];
	PlcInputs.ST80_1_DM260_PB_Box_Result_Data_64_bytes_1[40] := HwInputs.ST80_1_DM260_PB_Box_Result_Data_64_bytes_1[40];
	PlcInputs.ST80_1_DM260_PB_Box_Result_Data_64_bytes_1[41] := HwInputs.ST80_1_DM260_PB_Box_Result_Data_64_bytes_1[41];
	PlcInputs.ST80_1_DM260_PB_Box_Result_Data_64_bytes_1[42] := HwInputs.ST80_1_DM260_PB_Box_Result_Data_64_bytes_1[42];
	PlcInputs.ST80_1_DM260_PB_Box_Result_Data_64_bytes_1[43] := HwInputs.ST80_1_DM260_PB_Box_Result_Data_64_bytes_1[43];
	PlcInputs.ST80_1_DM260_PB_Box_Result_Data_64_bytes_1[44] := HwInputs.ST80_1_DM260_PB_Box_Result_Data_64_bytes_1[44];
	PlcInputs.ST80_1_DM260_PB_Box_Result_Data_64_bytes_1[45] := HwInputs.ST80_1_DM260_PB_Box_Result_Data_64_bytes_1[45];
	PlcInputs.ST80_1_DM260_PB_Box_Result_Data_64_bytes_1[46] := HwInputs.ST80_1_DM260_PB_Box_Result_Data_64_bytes_1[46];
	PlcInputs.ST80_1_DM260_PB_Box_Result_Data_64_bytes_1[47] := HwInputs.ST80_1_DM260_PB_Box_Result_Data_64_bytes_1[47];
	PlcInputs.ST80_1_DM260_PB_Box_Result_Data_64_bytes_1[48] := HwInputs.ST80_1_DM260_PB_Box_Result_Data_64_bytes_1[48];
	PlcInputs.ST80_1_DM260_PB_Box_Result_Data_64_bytes_1[49] := HwInputs.ST80_1_DM260_PB_Box_Result_Data_64_bytes_1[49];
	PlcInputs.ST80_1_DM260_PB_Box_Result_Data_64_bytes_1[50] := HwInputs.ST80_1_DM260_PB_Box_Result_Data_64_bytes_1[50];
	PlcInputs.ST80_1_DM260_PB_Box_Result_Data_64_bytes_1[51] := HwInputs.ST80_1_DM260_PB_Box_Result_Data_64_bytes_1[51];
	PlcInputs.ST80_1_DM260_PB_Box_Result_Data_64_bytes_1[52] := HwInputs.ST80_1_DM260_PB_Box_Result_Data_64_bytes_1[52];
	PlcInputs.ST80_1_DM260_PB_Box_Result_Data_64_bytes_1[53] := HwInputs.ST80_1_DM260_PB_Box_Result_Data_64_bytes_1[53];
	PlcInputs.ST80_1_DM260_PB_Box_Result_Data_64_bytes_1[54] := HwInputs.ST80_1_DM260_PB_Box_Result_Data_64_bytes_1[54];
	PlcInputs.ST80_1_DM260_PB_Box_Result_Data_64_bytes_1[55] := HwInputs.ST80_1_DM260_PB_Box_Result_Data_64_bytes_1[55];
	PlcInputs.ST80_1_DM260_PB_Box_Result_Data_64_bytes_1[56] := HwInputs.ST80_1_DM260_PB_Box_Result_Data_64_bytes_1[56];
	PlcInputs.ST80_1_DM260_PB_Box_Result_Data_64_bytes_1[57] := HwInputs.ST80_1_DM260_PB_Box_Result_Data_64_bytes_1[57];
	PlcInputs.ST80_1_DM260_PB_Box_Result_Data_64_bytes_1[58] := HwInputs.ST80_1_DM260_PB_Box_Result_Data_64_bytes_1[58];
	PlcInputs.ST80_1_DM260_PB_Box_Result_Data_64_bytes_1[59] := HwInputs.ST80_1_DM260_PB_Box_Result_Data_64_bytes_1[59];
	PlcInputs.ST80_1_DM260_PB_Box_Result_Data_64_bytes_1[60] := HwInputs.ST80_1_DM260_PB_Box_Result_Data_64_bytes_1[60];
	PlcInputs.ST80_1_DM260_PB_Box_Result_Data_64_bytes_1[61] := HwInputs.ST80_1_DM260_PB_Box_Result_Data_64_bytes_1[61];
	PlcInputs.ST80_1_DM260_PB_Box_Result_Data_64_bytes_1[62] := HwInputs.ST80_1_DM260_PB_Box_Result_Data_64_bytes_1[62];
	PlcInputs.ST80_1_DM260_PB_Box_Result_Data_64_bytes_1[63] := HwInputs.ST80_1_DM260_PB_Box_Result_Data_64_bytes_1[63];
	PlcInputs.ST80_1_DM260_PB_Box_Result_Data_64_bytes_1[64] := HwInputs.ST80_1_DM260_PB_Box_Result_Data_64_bytes_1[64];
	PlcInputs.ST80_1_DM260_PB_Box_Result_Data_64_bytes_1[65] := HwInputs.ST80_1_DM260_PB_Box_Result_Data_64_bytes_1[65];
	PlcInputs.ST80_1_DM260_PB_Box_Result_Data_64_bytes_1[66] := HwInputs.ST80_1_DM260_PB_Box_Result_Data_64_bytes_1[66];
	PlcInputs.ST80_1_DM260_PB_Box_Result_Data_64_bytes_1[67] := HwInputs.ST80_1_DM260_PB_Box_Result_Data_64_bytes_1[67];
	PlcInputs.ST80_1_DM260_PB_Box_Result_Data_64_bytes_1[68] := HwInputs.ST80_1_DM260_PB_Box_Result_Data_64_bytes_1[68];
	PlcInputs.ST80_1_DM260_PB_Box_Result_Data_64_bytes_1[69] := HwInputs.ST80_1_DM260_PB_Box_Result_Data_64_bytes_1[69];
	PlcInputs.ST80_1_DM260_PB_Box_Result_Data_64_bytes_1[70] := HwInputs.ST80_1_DM260_PB_Box_Result_Data_64_bytes_1[70];
	PlcInputs.ST80_1_DM260_PB_Box_Result_Data_64_bytes_1[71] := HwInputs.ST80_1_DM260_PB_Box_Result_Data_64_bytes_1[71];
	PlcInputs.ST80_ET200SP_2_11M1 := HwInputs.ST80_ET200SP_2_11M1;
	PlcInputs.ST80_ET200SP_2_11M2 := HwInputs.ST80_ET200SP_2_11M2;
	PlcInputs.ST80_ET200SP_2_11M3 := HwInputs.ST80_ET200SP_2_11M3;
	PlcInputs.ST80_ET200SP_2_11M4 := HwInputs.ST80_ET200SP_2_11M4;
	PlcInputs.ST80_ET200SP_2_12M1 := HwInputs.ST80_ET200SP_2_12M1;
	PlcInputs.ST80_ET200SP_2_12M2 := HwInputs.ST80_ET200SP_2_12M2;
	PlcInputs.ST80_ET200SP_2_12M3 := HwInputs.ST80_ET200SP_2_12M3;
	PlcInputs.ST80_ET200SP_2_12M4 := HwInputs.ST80_ET200SP_2_12M4;
	PlcInputs.ST80_ET200SP_2_13M1 := HwInputs.ST80_ET200SP_2_13M1;
	PlcInputs.ST80_ET200SP_2_13M2 := HwInputs.ST80_ET200SP_2_13M2;
	PlcInputs.ST80_ET200SP_2_13M3 := HwInputs.ST80_ET200SP_2_13M3;
	PlcInputs.ST80_ET200SP_2_13M4 := HwInputs.ST80_ET200SP_2_13M4;
	PlcInputs.ST80_1_TZ535_PN_In_Out_32_byte_1[0] := HwInputs.ST80_1_TZ535_PN_In_Out_32_byte_1[0];
	PlcInputs.ST80_1_TZ535_PN_In_Out_32_byte_1[1] := HwInputs.ST80_1_TZ535_PN_In_Out_32_byte_1[1];
	PlcInputs.ST80_1_TZ535_PN_In_Out_32_byte_1[2] := HwInputs.ST80_1_TZ535_PN_In_Out_32_byte_1[2];
	PlcInputs.ST80_1_TZ535_PN_In_Out_32_byte_1[3] := HwInputs.ST80_1_TZ535_PN_In_Out_32_byte_1[3];
	PlcInputs.ST80_1_TZ535_PN_In_Out_32_byte_1[4] := HwInputs.ST80_1_TZ535_PN_In_Out_32_byte_1[4];
	PlcInputs.ST80_1_TZ535_PN_In_Out_32_byte_1[5] := HwInputs.ST80_1_TZ535_PN_In_Out_32_byte_1[5];
	PlcInputs.ST80_1_TZ535_PN_In_Out_32_byte_1[6] := HwInputs.ST80_1_TZ535_PN_In_Out_32_byte_1[6];
	PlcInputs.ST80_1_TZ535_PN_In_Out_32_byte_1[7] := HwInputs.ST80_1_TZ535_PN_In_Out_32_byte_1[7];
	PlcInputs.ST80_1_TZ535_PN_In_Out_32_byte_1[8] := HwInputs.ST80_1_TZ535_PN_In_Out_32_byte_1[8];
	PlcInputs.ST80_1_TZ535_PN_In_Out_32_byte_1[9] := HwInputs.ST80_1_TZ535_PN_In_Out_32_byte_1[9];
	PlcInputs.ST80_1_TZ535_PN_In_Out_32_byte_1[10] := HwInputs.ST80_1_TZ535_PN_In_Out_32_byte_1[10];
	PlcInputs.ST80_1_TZ535_PN_In_Out_32_byte_1[11] := HwInputs.ST80_1_TZ535_PN_In_Out_32_byte_1[11];
	PlcInputs.ST80_1_TZ535_PN_In_Out_32_byte_1[12] := HwInputs.ST80_1_TZ535_PN_In_Out_32_byte_1[12];
	PlcInputs.ST80_1_TZ535_PN_In_Out_32_byte_1[13] := HwInputs.ST80_1_TZ535_PN_In_Out_32_byte_1[13];
	PlcInputs.ST80_1_TZ535_PN_In_Out_32_byte_1[14] := HwInputs.ST80_1_TZ535_PN_In_Out_32_byte_1[14];
	PlcInputs.ST80_1_TZ535_PN_In_Out_32_byte_1[15] := HwInputs.ST80_1_TZ535_PN_In_Out_32_byte_1[15];
	PlcInputs.ST80_1_TZ535_PN_In_Out_32_byte_1[16] := HwInputs.ST80_1_TZ535_PN_In_Out_32_byte_1[16];
	PlcInputs.ST80_1_TZ535_PN_In_Out_32_byte_1[17] := HwInputs.ST80_1_TZ535_PN_In_Out_32_byte_1[17];
	PlcInputs.ST80_1_TZ535_PN_In_Out_32_byte_1[18] := HwInputs.ST80_1_TZ535_PN_In_Out_32_byte_1[18];
	PlcInputs.ST80_1_TZ535_PN_In_Out_32_byte_1[19] := HwInputs.ST80_1_TZ535_PN_In_Out_32_byte_1[19];
	PlcInputs.ST80_1_TZ535_PN_In_Out_32_byte_1[20] := HwInputs.ST80_1_TZ535_PN_In_Out_32_byte_1[20];
	PlcInputs.ST80_1_TZ535_PN_In_Out_32_byte_1[21] := HwInputs.ST80_1_TZ535_PN_In_Out_32_byte_1[21];
	PlcInputs.ST80_1_TZ535_PN_In_Out_32_byte_1[22] := HwInputs.ST80_1_TZ535_PN_In_Out_32_byte_1[22];
	PlcInputs.ST80_1_TZ535_PN_In_Out_32_byte_1[23] := HwInputs.ST80_1_TZ535_PN_In_Out_32_byte_1[23];
	PlcInputs.ST80_1_TZ535_PN_In_Out_32_byte_1[24] := HwInputs.ST80_1_TZ535_PN_In_Out_32_byte_1[24];
	PlcInputs.ST80_1_TZ535_PN_In_Out_32_byte_1[25] := HwInputs.ST80_1_TZ535_PN_In_Out_32_byte_1[25];
	PlcInputs.ST80_1_TZ535_PN_In_Out_32_byte_1[26] := HwInputs.ST80_1_TZ535_PN_In_Out_32_byte_1[26];
	PlcInputs.ST80_1_TZ535_PN_In_Out_32_byte_1[27] := HwInputs.ST80_1_TZ535_PN_In_Out_32_byte_1[27];
	PlcInputs.ST80_1_TZ535_PN_In_Out_32_byte_1[28] := HwInputs.ST80_1_TZ535_PN_In_Out_32_byte_1[28];
	PlcInputs.ST80_1_TZ535_PN_In_Out_32_byte_1[29] := HwInputs.ST80_1_TZ535_PN_In_Out_32_byte_1[29];
	PlcInputs.ST80_1_TZ535_PN_In_Out_32_byte_1[30] := HwInputs.ST80_1_TZ535_PN_In_Out_32_byte_1[30];
	PlcInputs.ST80_1_TZ535_PN_In_Out_32_byte_1[31] := HwInputs.ST80_1_TZ535_PN_In_Out_32_byte_1[31];
	PlcInputs.ST80_1_DM260_Housing_Acquisition_Status_1[0] := HwInputs.ST80_1_DM260_Housing_Acquisition_Status_1[0];
	PlcInputs.ST80_1_DM260_Housing_Acquisition_Status_1[1] := HwInputs.ST80_1_DM260_Housing_Acquisition_Status_1[1];
	PlcInputs.ST80_1_DM260_Housing_Acquisition_Status_1[2] := HwInputs.ST80_1_DM260_Housing_Acquisition_Status_1[2];
	PlcInputs.ST80_1_DM260_Housing_Results_Status_1 := HwInputs.ST80_1_DM260_Housing_Results_Status_1;
	PlcInputs.ST80_1_DM260_Housing_Soft_Event_Control_1 := HwInputs.ST80_1_DM260_Housing_Soft_Event_Control_1;
	PlcInputs.ST80_1_DM260_Housing_Result_Data_64_bytes_1[0] := HwInputs.ST80_1_DM260_Housing_Result_Data_64_bytes_1[0];
	PlcInputs.ST80_1_DM260_Housing_Result_Data_64_bytes_1[1] := HwInputs.ST80_1_DM260_Housing_Result_Data_64_bytes_1[1];
	PlcInputs.ST80_1_DM260_Housing_Result_Data_64_bytes_1[2] := HwInputs.ST80_1_DM260_Housing_Result_Data_64_bytes_1[2];
	PlcInputs.ST80_1_DM260_Housing_Result_Data_64_bytes_1[3] := HwInputs.ST80_1_DM260_Housing_Result_Data_64_bytes_1[3];
	PlcInputs.ST80_1_DM260_Housing_Result_Data_64_bytes_1[4] := HwInputs.ST80_1_DM260_Housing_Result_Data_64_bytes_1[4];
	PlcInputs.ST80_1_DM260_Housing_Result_Data_64_bytes_1[5] := HwInputs.ST80_1_DM260_Housing_Result_Data_64_bytes_1[5];
	PlcInputs.ST80_1_DM260_Housing_Result_Data_64_bytes_1[6] := HwInputs.ST80_1_DM260_Housing_Result_Data_64_bytes_1[6];
	PlcInputs.ST80_1_DM260_Housing_Result_Data_64_bytes_1[7] := HwInputs.ST80_1_DM260_Housing_Result_Data_64_bytes_1[7];
	PlcInputs.ST80_1_DM260_Housing_Result_Data_64_bytes_1[8] := HwInputs.ST80_1_DM260_Housing_Result_Data_64_bytes_1[8];
	PlcInputs.ST80_1_DM260_Housing_Result_Data_64_bytes_1[9] := HwInputs.ST80_1_DM260_Housing_Result_Data_64_bytes_1[9];
	PlcInputs.ST80_1_DM260_Housing_Result_Data_64_bytes_1[10] := HwInputs.ST80_1_DM260_Housing_Result_Data_64_bytes_1[10];
	PlcInputs.ST80_1_DM260_Housing_Result_Data_64_bytes_1[11] := HwInputs.ST80_1_DM260_Housing_Result_Data_64_bytes_1[11];
	PlcInputs.ST80_1_DM260_Housing_Result_Data_64_bytes_1[12] := HwInputs.ST80_1_DM260_Housing_Result_Data_64_bytes_1[12];
	PlcInputs.ST80_1_DM260_Housing_Result_Data_64_bytes_1[13] := HwInputs.ST80_1_DM260_Housing_Result_Data_64_bytes_1[13];
	PlcInputs.ST80_1_DM260_Housing_Result_Data_64_bytes_1[14] := HwInputs.ST80_1_DM260_Housing_Result_Data_64_bytes_1[14];
	PlcInputs.ST80_1_DM260_Housing_Result_Data_64_bytes_1[15] := HwInputs.ST80_1_DM260_Housing_Result_Data_64_bytes_1[15];
	PlcInputs.ST80_1_DM260_Housing_Result_Data_64_bytes_1[16] := HwInputs.ST80_1_DM260_Housing_Result_Data_64_bytes_1[16];
	PlcInputs.ST80_1_DM260_Housing_Result_Data_64_bytes_1[17] := HwInputs.ST80_1_DM260_Housing_Result_Data_64_bytes_1[17];
	PlcInputs.ST80_1_DM260_Housing_Result_Data_64_bytes_1[18] := HwInputs.ST80_1_DM260_Housing_Result_Data_64_bytes_1[18];
	PlcInputs.ST80_1_DM260_Housing_Result_Data_64_bytes_1[19] := HwInputs.ST80_1_DM260_Housing_Result_Data_64_bytes_1[19];
	PlcInputs.ST80_1_DM260_Housing_Result_Data_64_bytes_1[20] := HwInputs.ST80_1_DM260_Housing_Result_Data_64_bytes_1[20];
	PlcInputs.ST80_1_DM260_Housing_Result_Data_64_bytes_1[21] := HwInputs.ST80_1_DM260_Housing_Result_Data_64_bytes_1[21];
	PlcInputs.ST80_1_DM260_Housing_Result_Data_64_bytes_1[22] := HwInputs.ST80_1_DM260_Housing_Result_Data_64_bytes_1[22];
	PlcInputs.ST80_1_DM260_Housing_Result_Data_64_bytes_1[23] := HwInputs.ST80_1_DM260_Housing_Result_Data_64_bytes_1[23];
	PlcInputs.ST80_1_DM260_Housing_Result_Data_64_bytes_1[24] := HwInputs.ST80_1_DM260_Housing_Result_Data_64_bytes_1[24];
	PlcInputs.ST80_1_DM260_Housing_Result_Data_64_bytes_1[25] := HwInputs.ST80_1_DM260_Housing_Result_Data_64_bytes_1[25];
	PlcInputs.ST80_1_DM260_Housing_Result_Data_64_bytes_1[26] := HwInputs.ST80_1_DM260_Housing_Result_Data_64_bytes_1[26];
	PlcInputs.ST80_1_DM260_Housing_Result_Data_64_bytes_1[27] := HwInputs.ST80_1_DM260_Housing_Result_Data_64_bytes_1[27];
	PlcInputs.ST80_1_DM260_Housing_Result_Data_64_bytes_1[28] := HwInputs.ST80_1_DM260_Housing_Result_Data_64_bytes_1[28];
	PlcInputs.ST80_1_DM260_Housing_Result_Data_64_bytes_1[29] := HwInputs.ST80_1_DM260_Housing_Result_Data_64_bytes_1[29];
	PlcInputs.ST80_1_DM260_Housing_Result_Data_64_bytes_1[30] := HwInputs.ST80_1_DM260_Housing_Result_Data_64_bytes_1[30];
	PlcInputs.ST80_1_DM260_Housing_Result_Data_64_bytes_1[31] := HwInputs.ST80_1_DM260_Housing_Result_Data_64_bytes_1[31];
	PlcInputs.ST80_1_DM260_Housing_Result_Data_64_bytes_1[32] := HwInputs.ST80_1_DM260_Housing_Result_Data_64_bytes_1[32];
	PlcInputs.ST80_1_DM260_Housing_Result_Data_64_bytes_1[33] := HwInputs.ST80_1_DM260_Housing_Result_Data_64_bytes_1[33];
	PlcInputs.ST80_1_DM260_Housing_Result_Data_64_bytes_1[34] := HwInputs.ST80_1_DM260_Housing_Result_Data_64_bytes_1[34];
	PlcInputs.ST80_1_DM260_Housing_Result_Data_64_bytes_1[35] := HwInputs.ST80_1_DM260_Housing_Result_Data_64_bytes_1[35];
	PlcInputs.ST80_1_DM260_Housing_Result_Data_64_bytes_1[36] := HwInputs.ST80_1_DM260_Housing_Result_Data_64_bytes_1[36];
	PlcInputs.ST80_1_DM260_Housing_Result_Data_64_bytes_1[37] := HwInputs.ST80_1_DM260_Housing_Result_Data_64_bytes_1[37];
	PlcInputs.ST80_1_DM260_Housing_Result_Data_64_bytes_1[38] := HwInputs.ST80_1_DM260_Housing_Result_Data_64_bytes_1[38];
	PlcInputs.ST80_1_DM260_Housing_Result_Data_64_bytes_1[39] := HwInputs.ST80_1_DM260_Housing_Result_Data_64_bytes_1[39];
	PlcInputs.ST80_1_DM260_Housing_Result_Data_64_bytes_1[40] := HwInputs.ST80_1_DM260_Housing_Result_Data_64_bytes_1[40];
	PlcInputs.ST80_1_DM260_Housing_Result_Data_64_bytes_1[41] := HwInputs.ST80_1_DM260_Housing_Result_Data_64_bytes_1[41];
	PlcInputs.ST80_1_DM260_Housing_Result_Data_64_bytes_1[42] := HwInputs.ST80_1_DM260_Housing_Result_Data_64_bytes_1[42];
	PlcInputs.ST80_1_DM260_Housing_Result_Data_64_bytes_1[43] := HwInputs.ST80_1_DM260_Housing_Result_Data_64_bytes_1[43];
	PlcInputs.ST80_1_DM260_Housing_Result_Data_64_bytes_1[44] := HwInputs.ST80_1_DM260_Housing_Result_Data_64_bytes_1[44];
	PlcInputs.ST80_1_DM260_Housing_Result_Data_64_bytes_1[45] := HwInputs.ST80_1_DM260_Housing_Result_Data_64_bytes_1[45];
	PlcInputs.ST80_1_DM260_Housing_Result_Data_64_bytes_1[46] := HwInputs.ST80_1_DM260_Housing_Result_Data_64_bytes_1[46];
	PlcInputs.ST80_1_DM260_Housing_Result_Data_64_bytes_1[47] := HwInputs.ST80_1_DM260_Housing_Result_Data_64_bytes_1[47];
	PlcInputs.ST80_1_DM260_Housing_Result_Data_64_bytes_1[48] := HwInputs.ST80_1_DM260_Housing_Result_Data_64_bytes_1[48];
	PlcInputs.ST80_1_DM260_Housing_Result_Data_64_bytes_1[49] := HwInputs.ST80_1_DM260_Housing_Result_Data_64_bytes_1[49];
	PlcInputs.ST80_1_DM260_Housing_Result_Data_64_bytes_1[50] := HwInputs.ST80_1_DM260_Housing_Result_Data_64_bytes_1[50];
	PlcInputs.ST80_1_DM260_Housing_Result_Data_64_bytes_1[51] := HwInputs.ST80_1_DM260_Housing_Result_Data_64_bytes_1[51];
	PlcInputs.ST80_1_DM260_Housing_Result_Data_64_bytes_1[52] := HwInputs.ST80_1_DM260_Housing_Result_Data_64_bytes_1[52];
	PlcInputs.ST80_1_DM260_Housing_Result_Data_64_bytes_1[53] := HwInputs.ST80_1_DM260_Housing_Result_Data_64_bytes_1[53];
	PlcInputs.ST80_1_DM260_Housing_Result_Data_64_bytes_1[54] := HwInputs.ST80_1_DM260_Housing_Result_Data_64_bytes_1[54];
	PlcInputs.ST80_1_DM260_Housing_Result_Data_64_bytes_1[55] := HwInputs.ST80_1_DM260_Housing_Result_Data_64_bytes_1[55];
	PlcInputs.ST80_1_DM260_Housing_Result_Data_64_bytes_1[56] := HwInputs.ST80_1_DM260_Housing_Result_Data_64_bytes_1[56];
	PlcInputs.ST80_1_DM260_Housing_Result_Data_64_bytes_1[57] := HwInputs.ST80_1_DM260_Housing_Result_Data_64_bytes_1[57];
	PlcInputs.ST80_1_DM260_Housing_Result_Data_64_bytes_1[58] := HwInputs.ST80_1_DM260_Housing_Result_Data_64_bytes_1[58];
	PlcInputs.ST80_1_DM260_Housing_Result_Data_64_bytes_1[59] := HwInputs.ST80_1_DM260_Housing_Result_Data_64_bytes_1[59];
	PlcInputs.ST80_1_DM260_Housing_Result_Data_64_bytes_1[60] := HwInputs.ST80_1_DM260_Housing_Result_Data_64_bytes_1[60];
	PlcInputs.ST80_1_DM260_Housing_Result_Data_64_bytes_1[61] := HwInputs.ST80_1_DM260_Housing_Result_Data_64_bytes_1[61];
	PlcInputs.ST80_1_DM260_Housing_Result_Data_64_bytes_1[62] := HwInputs.ST80_1_DM260_Housing_Result_Data_64_bytes_1[62];
	PlcInputs.ST80_1_DM260_Housing_Result_Data_64_bytes_1[63] := HwInputs.ST80_1_DM260_Housing_Result_Data_64_bytes_1[63];
	PlcInputs.ST80_1_DM260_Housing_Result_Data_64_bytes_1[64] := HwInputs.ST80_1_DM260_Housing_Result_Data_64_bytes_1[64];
	PlcInputs.ST80_1_DM260_Housing_Result_Data_64_bytes_1[65] := HwInputs.ST80_1_DM260_Housing_Result_Data_64_bytes_1[65];
	PlcInputs.ST80_1_DM260_Housing_Result_Data_64_bytes_1[66] := HwInputs.ST80_1_DM260_Housing_Result_Data_64_bytes_1[66];
	PlcInputs.ST80_1_DM260_Housing_Result_Data_64_bytes_1[67] := HwInputs.ST80_1_DM260_Housing_Result_Data_64_bytes_1[67];
	PlcInputs.ST80_1_DM260_Housing_Result_Data_64_bytes_1[68] := HwInputs.ST80_1_DM260_Housing_Result_Data_64_bytes_1[68];
	PlcInputs.ST80_1_DM260_Housing_Result_Data_64_bytes_1[69] := HwInputs.ST80_1_DM260_Housing_Result_Data_64_bytes_1[69];
	PlcInputs.ST80_1_DM260_Housing_Result_Data_64_bytes_1[70] := HwInputs.ST80_1_DM260_Housing_Result_Data_64_bytes_1[70];
	PlcInputs.ST80_1_DM260_Housing_Result_Data_64_bytes_1[71] := HwInputs.ST80_1_DM260_Housing_Result_Data_64_bytes_1[71];
	PlcInputs.ST80_1_CMMT_3GF1_DO_SERVO_1_Siemens_telegram_111_PZD_12_12[0] := HwInputs.ST80_1_CMMT_3GF1_DO_SERVO_1_Siemens_telegram_111_PZD_12_12[0];
	PlcInputs.ST80_1_CMMT_3GF1_DO_SERVO_1_Siemens_telegram_111_PZD_12_12[1] := HwInputs.ST80_1_CMMT_3GF1_DO_SERVO_1_Siemens_telegram_111_PZD_12_12[1];
	PlcInputs.ST80_1_CMMT_3GF1_DO_SERVO_1_Siemens_telegram_111_PZD_12_12[2] := HwInputs.ST80_1_CMMT_3GF1_DO_SERVO_1_Siemens_telegram_111_PZD_12_12[2];
	PlcInputs.ST80_1_CMMT_3GF1_DO_SERVO_1_Siemens_telegram_111_PZD_12_12[3] := HwInputs.ST80_1_CMMT_3GF1_DO_SERVO_1_Siemens_telegram_111_PZD_12_12[3];
	PlcInputs.ST80_1_CMMT_3GF1_DO_SERVO_1_Siemens_telegram_111_PZD_12_12[4] := HwInputs.ST80_1_CMMT_3GF1_DO_SERVO_1_Siemens_telegram_111_PZD_12_12[4];
	PlcInputs.ST80_1_CMMT_3GF1_DO_SERVO_1_Siemens_telegram_111_PZD_12_12[5] := HwInputs.ST80_1_CMMT_3GF1_DO_SERVO_1_Siemens_telegram_111_PZD_12_12[5];
	PlcInputs.ST80_1_CMMT_3GF1_DO_SERVO_1_Siemens_telegram_111_PZD_12_12[6] := HwInputs.ST80_1_CMMT_3GF1_DO_SERVO_1_Siemens_telegram_111_PZD_12_12[6];
	PlcInputs.ST80_1_CMMT_3GF1_DO_SERVO_1_Siemens_telegram_111_PZD_12_12[7] := HwInputs.ST80_1_CMMT_3GF1_DO_SERVO_1_Siemens_telegram_111_PZD_12_12[7];
	PlcInputs.ST80_1_CMMT_3GF1_DO_SERVO_1_Siemens_telegram_111_PZD_12_12[8] := HwInputs.ST80_1_CMMT_3GF1_DO_SERVO_1_Siemens_telegram_111_PZD_12_12[8];
	PlcInputs.ST80_1_CMMT_3GF1_DO_SERVO_1_Siemens_telegram_111_PZD_12_12[9] := HwInputs.ST80_1_CMMT_3GF1_DO_SERVO_1_Siemens_telegram_111_PZD_12_12[9];
	PlcInputs.ST80_1_CMMT_3GF1_DO_SERVO_1_Siemens_telegram_111_PZD_12_12[10] := HwInputs.ST80_1_CMMT_3GF1_DO_SERVO_1_Siemens_telegram_111_PZD_12_12[10];
	PlcInputs.ST80_1_CMMT_3GF1_DO_SERVO_1_Siemens_telegram_111_PZD_12_12[11] := HwInputs.ST80_1_CMMT_3GF1_DO_SERVO_1_Siemens_telegram_111_PZD_12_12[11];
	PlcInputs.ST80_1_CMMT_3GF1_DO_SERVO_1_Siemens_telegram_111_PZD_12_12[12] := HwInputs.ST80_1_CMMT_3GF1_DO_SERVO_1_Siemens_telegram_111_PZD_12_12[12];
	PlcInputs.ST80_1_CMMT_3GF1_DO_SERVO_1_Siemens_telegram_111_PZD_12_12[13] := HwInputs.ST80_1_CMMT_3GF1_DO_SERVO_1_Siemens_telegram_111_PZD_12_12[13];
	PlcInputs.ST80_1_CMMT_3GF1_DO_SERVO_1_Siemens_telegram_111_PZD_12_12[14] := HwInputs.ST80_1_CMMT_3GF1_DO_SERVO_1_Siemens_telegram_111_PZD_12_12[14];
	PlcInputs.ST80_1_CMMT_3GF1_DO_SERVO_1_Siemens_telegram_111_PZD_12_12[15] := HwInputs.ST80_1_CMMT_3GF1_DO_SERVO_1_Siemens_telegram_111_PZD_12_12[15];
	PlcInputs.ST80_1_CMMT_3GF1_DO_SERVO_1_Siemens_telegram_111_PZD_12_12[16] := HwInputs.ST80_1_CMMT_3GF1_DO_SERVO_1_Siemens_telegram_111_PZD_12_12[16];
	PlcInputs.ST80_1_CMMT_3GF1_DO_SERVO_1_Siemens_telegram_111_PZD_12_12[17] := HwInputs.ST80_1_CMMT_3GF1_DO_SERVO_1_Siemens_telegram_111_PZD_12_12[17];
	PlcInputs.ST80_1_CMMT_3GF1_DO_SERVO_1_Siemens_telegram_111_PZD_12_12[18] := HwInputs.ST80_1_CMMT_3GF1_DO_SERVO_1_Siemens_telegram_111_PZD_12_12[18];
	PlcInputs.ST80_1_CMMT_3GF1_DO_SERVO_1_Siemens_telegram_111_PZD_12_12[19] := HwInputs.ST80_1_CMMT_3GF1_DO_SERVO_1_Siemens_telegram_111_PZD_12_12[19];
	PlcInputs.ST80_1_CMMT_3GF1_DO_SERVO_1_Siemens_telegram_111_PZD_12_12[20] := HwInputs.ST80_1_CMMT_3GF1_DO_SERVO_1_Siemens_telegram_111_PZD_12_12[20];
	PlcInputs.ST80_1_CMMT_3GF1_DO_SERVO_1_Siemens_telegram_111_PZD_12_12[21] := HwInputs.ST80_1_CMMT_3GF1_DO_SERVO_1_Siemens_telegram_111_PZD_12_12[21];
	PlcInputs.ST80_1_CMMT_3GF1_DO_SERVO_1_Siemens_telegram_111_PZD_12_12[22] := HwInputs.ST80_1_CMMT_3GF1_DO_SERVO_1_Siemens_telegram_111_PZD_12_12[22];
	PlcInputs.ST80_1_CMMT_3GF1_DO_SERVO_1_Siemens_telegram_111_PZD_12_12[23] := HwInputs.ST80_1_CMMT_3GF1_DO_SERVO_1_Siemens_telegram_111_PZD_12_12[23];
	PlcInputs.ST80_ET200SP_CM_4xIO_Link_1[0] := HwInputs.ST80_ET200SP_CM_4xIO_Link_1[0];
	PlcInputs.ST80_ET200SP_CM_4xIO_Link_1[1] := HwInputs.ST80_ET200SP_CM_4xIO_Link_1[1];
	PlcInputs.ST80_ET200SP_CM_4xIO_Link_1[2] := HwInputs.ST80_ET200SP_CM_4xIO_Link_1[2];
	PlcInputs.ST80_ET200SP_CM_4xIO_Link_1[3] := HwInputs.ST80_ET200SP_CM_4xIO_Link_1[3];
	PlcInputs.ST80_ET200SP_CM_4xIO_Link_1[4] := HwInputs.ST80_ET200SP_CM_4xIO_Link_1[4];
	PlcInputs.ST80_ET200SP_CM_4xIO_Link_1[5] := HwInputs.ST80_ET200SP_CM_4xIO_Link_1[5];
	PlcInputs.ST80_ET200SP_CM_4xIO_Link_1[6] := HwInputs.ST80_ET200SP_CM_4xIO_Link_1[6];
	PlcInputs.ST80_ET200SP_CM_4xIO_Link_1[7] := HwInputs.ST80_ET200SP_CM_4xIO_Link_1[7];
	PlcInputs.ST80_ET200SP_CM_4xIO_Link_1[8] := HwInputs.ST80_ET200SP_CM_4xIO_Link_1[8];
	PlcInputs.ST80_ET200SP_CM_4xIO_Link_1[9] := HwInputs.ST80_ET200SP_CM_4xIO_Link_1[9];
	PlcInputs.ST80_ET200SP_CM_4xIO_Link_1[10] := HwInputs.ST80_ET200SP_CM_4xIO_Link_1[10];
	PlcInputs.ST80_ET200SP_CM_4xIO_Link_1[11] := HwInputs.ST80_ET200SP_CM_4xIO_Link_1[11];
	PlcInputs.ST80_ET200SP_CM_4xIO_Link_1[12] := HwInputs.ST80_ET200SP_CM_4xIO_Link_1[12];
	PlcInputs.ST80_ET200SP_CM_4xIO_Link_1[13] := HwInputs.ST80_ET200SP_CM_4xIO_Link_1[13];
	PlcInputs.ST80_ET200SP_CM_4xIO_Link_1[14] := HwInputs.ST80_ET200SP_CM_4xIO_Link_1[14];
	PlcInputs.ST80_ET200SP_CM_4xIO_Link_1[15] := HwInputs.ST80_ET200SP_CM_4xIO_Link_1[15];
	PlcInputs.ST80_ET200SP_CM_4xIO_Link_1[16] := HwInputs.ST80_ET200SP_CM_4xIO_Link_1[16];
	PlcInputs.ST80_ET200SP_CM_4xIO_Link_1[17] := HwInputs.ST80_ET200SP_CM_4xIO_Link_1[17];
	PlcInputs.ST80_ET200SP_CM_4xIO_Link_1[18] := HwInputs.ST80_ET200SP_CM_4xIO_Link_1[18];
	PlcInputs.ST80_ET200SP_CM_4xIO_Link_1[19] := HwInputs.ST80_ET200SP_CM_4xIO_Link_1[19];
	PlcInputs.ST80_ET200SP_CM_4xIO_Link_1[20] := HwInputs.ST80_ET200SP_CM_4xIO_Link_1[20];
	PlcInputs.ST80_ET200SP_CM_4xIO_Link_1[21] := HwInputs.ST80_ET200SP_CM_4xIO_Link_1[21];
	PlcInputs.ST80_ET200SP_CM_4xIO_Link_1[22] := HwInputs.ST80_ET200SP_CM_4xIO_Link_1[22];
	PlcInputs.ST80_ET200SP_CM_4xIO_Link_1[23] := HwInputs.ST80_ET200SP_CM_4xIO_Link_1[23];
	PlcInputs.ST80_ET200SP_CM_4xIO_Link_1[24] := HwInputs.ST80_ET200SP_CM_4xIO_Link_1[24];
	PlcInputs.ST80_ET200SP_CM_4xIO_Link_1[25] := HwInputs.ST80_ET200SP_CM_4xIO_Link_1[25];
	PlcInputs.ST80_ET200SP_CM_4xIO_Link_1[26] := HwInputs.ST80_ET200SP_CM_4xIO_Link_1[26];
	PlcInputs.ST80_ET200SP_CM_4xIO_Link_1[27] := HwInputs.ST80_ET200SP_CM_4xIO_Link_1[27];
	PlcInputs.ST80_ET200SP_CM_4xIO_Link_1[28] := HwInputs.ST80_ET200SP_CM_4xIO_Link_1[28];
	PlcInputs.ST80_ET200SP_CM_4xIO_Link_1[29] := HwInputs.ST80_ET200SP_CM_4xIO_Link_1[29];
	PlcInputs.ST80_ET200SP_CM_4xIO_Link_1[30] := HwInputs.ST80_ET200SP_CM_4xIO_Link_1[30];
	PlcInputs.ST80_ET200SP_CM_4xIO_Link_1[31] := HwInputs.ST80_ET200SP_CM_4xIO_Link_1[31];
	PlcInputs.ST80_ET200SP_CM_4xIO_Link_2[0] := HwInputs.ST80_ET200SP_CM_4xIO_Link_2[0];
	PlcInputs.ST80_ET200SP_CM_4xIO_Link_2[1] := HwInputs.ST80_ET200SP_CM_4xIO_Link_2[1];
	PlcInputs.ST80_ET200SP_CM_4xIO_Link_2[2] := HwInputs.ST80_ET200SP_CM_4xIO_Link_2[2];
	PlcInputs.ST80_ET200SP_CM_4xIO_Link_2[3] := HwInputs.ST80_ET200SP_CM_4xIO_Link_2[3];
	PlcInputs.ST80_ET200SP_CM_4xIO_Link_2[4] := HwInputs.ST80_ET200SP_CM_4xIO_Link_2[4];
	PlcInputs.ST80_ET200SP_CM_4xIO_Link_2[5] := HwInputs.ST80_ET200SP_CM_4xIO_Link_2[5];
	PlcInputs.ST80_ET200SP_CM_4xIO_Link_2[6] := HwInputs.ST80_ET200SP_CM_4xIO_Link_2[6];
	PlcInputs.ST80_ET200SP_CM_4xIO_Link_2[7] := HwInputs.ST80_ET200SP_CM_4xIO_Link_2[7];
	PlcInputs.ST80_ET200SP_CM_4xIO_Link_2[8] := HwInputs.ST80_ET200SP_CM_4xIO_Link_2[8];
	PlcInputs.ST80_ET200SP_CM_4xIO_Link_2[9] := HwInputs.ST80_ET200SP_CM_4xIO_Link_2[9];
	PlcInputs.ST80_ET200SP_CM_4xIO_Link_2[10] := HwInputs.ST80_ET200SP_CM_4xIO_Link_2[10];
	PlcInputs.ST80_ET200SP_CM_4xIO_Link_2[11] := HwInputs.ST80_ET200SP_CM_4xIO_Link_2[11];
	PlcInputs.ST80_ET200SP_CM_4xIO_Link_2[12] := HwInputs.ST80_ET200SP_CM_4xIO_Link_2[12];
	PlcInputs.ST80_ET200SP_CM_4xIO_Link_2[13] := HwInputs.ST80_ET200SP_CM_4xIO_Link_2[13];
	PlcInputs.ST80_ET200SP_CM_4xIO_Link_2[14] := HwInputs.ST80_ET200SP_CM_4xIO_Link_2[14];
	PlcInputs.ST80_ET200SP_CM_4xIO_Link_2[15] := HwInputs.ST80_ET200SP_CM_4xIO_Link_2[15];
	PlcInputs.ST80_ET200SP_CM_4xIO_Link_2[16] := HwInputs.ST80_ET200SP_CM_4xIO_Link_2[16];
	PlcInputs.ST80_ET200SP_CM_4xIO_Link_2[17] := HwInputs.ST80_ET200SP_CM_4xIO_Link_2[17];
	PlcInputs.ST80_ET200SP_CM_4xIO_Link_2[18] := HwInputs.ST80_ET200SP_CM_4xIO_Link_2[18];
	PlcInputs.ST80_ET200SP_CM_4xIO_Link_2[19] := HwInputs.ST80_ET200SP_CM_4xIO_Link_2[19];
	PlcInputs.ST80_ET200SP_CM_4xIO_Link_2[20] := HwInputs.ST80_ET200SP_CM_4xIO_Link_2[20];
	PlcInputs.ST80_ET200SP_CM_4xIO_Link_2[21] := HwInputs.ST80_ET200SP_CM_4xIO_Link_2[21];
	PlcInputs.ST80_ET200SP_CM_4xIO_Link_2[22] := HwInputs.ST80_ET200SP_CM_4xIO_Link_2[22];
	PlcInputs.ST80_ET200SP_CM_4xIO_Link_2[23] := HwInputs.ST80_ET200SP_CM_4xIO_Link_2[23];
	PlcInputs.ST80_ET200SP_CM_4xIO_Link_2[24] := HwInputs.ST80_ET200SP_CM_4xIO_Link_2[24];
	PlcInputs.ST80_ET200SP_CM_4xIO_Link_2[25] := HwInputs.ST80_ET200SP_CM_4xIO_Link_2[25];
	PlcInputs.ST80_ET200SP_CM_4xIO_Link_2[26] := HwInputs.ST80_ET200SP_CM_4xIO_Link_2[26];
	PlcInputs.ST80_ET200SP_CM_4xIO_Link_2[27] := HwInputs.ST80_ET200SP_CM_4xIO_Link_2[27];
	PlcInputs.ST80_ET200SP_CM_4xIO_Link_2[28] := HwInputs.ST80_ET200SP_CM_4xIO_Link_2[28];
	PlcInputs.ST80_ET200SP_CM_4xIO_Link_2[29] := HwInputs.ST80_ET200SP_CM_4xIO_Link_2[29];
	PlcInputs.ST80_ET200SP_CM_4xIO_Link_2[30] := HwInputs.ST80_ET200SP_CM_4xIO_Link_2[30];
	PlcInputs.ST80_ET200SP_CM_4xIO_Link_2[31] := HwInputs.ST80_ET200SP_CM_4xIO_Link_2[31];
	PlcInputs.ST80_ET200SP_CM_4xIO_Link_3[0] := HwInputs.ST80_ET200SP_CM_4xIO_Link_3[0];
	PlcInputs.ST80_ET200SP_CM_4xIO_Link_3[1] := HwInputs.ST80_ET200SP_CM_4xIO_Link_3[1];
	PlcInputs.ST80_ET200SP_CM_4xIO_Link_3[2] := HwInputs.ST80_ET200SP_CM_4xIO_Link_3[2];
	PlcInputs.ST80_ET200SP_CM_4xIO_Link_3[3] := HwInputs.ST80_ET200SP_CM_4xIO_Link_3[3];
	PlcInputs.ST80_ET200SP_CM_4xIO_Link_3[4] := HwInputs.ST80_ET200SP_CM_4xIO_Link_3[4];
	PlcInputs.ST80_ET200SP_CM_4xIO_Link_3[5] := HwInputs.ST80_ET200SP_CM_4xIO_Link_3[5];
	PlcInputs.ST80_ET200SP_CM_4xIO_Link_3[6] := HwInputs.ST80_ET200SP_CM_4xIO_Link_3[6];
	PlcInputs.ST80_ET200SP_CM_4xIO_Link_3[7] := HwInputs.ST80_ET200SP_CM_4xIO_Link_3[7];
	PlcInputs.ST80_ET200SP_CM_4xIO_Link_3[8] := HwInputs.ST80_ET200SP_CM_4xIO_Link_3[8];
	PlcInputs.ST80_ET200SP_CM_4xIO_Link_3[9] := HwInputs.ST80_ET200SP_CM_4xIO_Link_3[9];
	PlcInputs.ST80_ET200SP_CM_4xIO_Link_3[10] := HwInputs.ST80_ET200SP_CM_4xIO_Link_3[10];
	PlcInputs.ST80_ET200SP_CM_4xIO_Link_3[11] := HwInputs.ST80_ET200SP_CM_4xIO_Link_3[11];
	PlcInputs.ST80_ET200SP_CM_4xIO_Link_3[12] := HwInputs.ST80_ET200SP_CM_4xIO_Link_3[12];
	PlcInputs.ST80_ET200SP_CM_4xIO_Link_3[13] := HwInputs.ST80_ET200SP_CM_4xIO_Link_3[13];
	PlcInputs.ST80_ET200SP_CM_4xIO_Link_3[14] := HwInputs.ST80_ET200SP_CM_4xIO_Link_3[14];
	PlcInputs.ST80_ET200SP_CM_4xIO_Link_3[15] := HwInputs.ST80_ET200SP_CM_4xIO_Link_3[15];
	PlcInputs.ST80_ET200SP_CM_4xIO_Link_3[16] := HwInputs.ST80_ET200SP_CM_4xIO_Link_3[16];
	PlcInputs.ST80_ET200SP_CM_4xIO_Link_3[17] := HwInputs.ST80_ET200SP_CM_4xIO_Link_3[17];
	PlcInputs.ST80_ET200SP_CM_4xIO_Link_3[18] := HwInputs.ST80_ET200SP_CM_4xIO_Link_3[18];
	PlcInputs.ST80_ET200SP_CM_4xIO_Link_3[19] := HwInputs.ST80_ET200SP_CM_4xIO_Link_3[19];
	PlcInputs.ST80_ET200SP_CM_4xIO_Link_3[20] := HwInputs.ST80_ET200SP_CM_4xIO_Link_3[20];
	PlcInputs.ST80_ET200SP_CM_4xIO_Link_3[21] := HwInputs.ST80_ET200SP_CM_4xIO_Link_3[21];
	PlcInputs.ST80_ET200SP_CM_4xIO_Link_3[22] := HwInputs.ST80_ET200SP_CM_4xIO_Link_3[22];
	PlcInputs.ST80_ET200SP_CM_4xIO_Link_3[23] := HwInputs.ST80_ET200SP_CM_4xIO_Link_3[23];
	PlcInputs.ST80_ET200SP_CM_4xIO_Link_3[24] := HwInputs.ST80_ET200SP_CM_4xIO_Link_3[24];
	PlcInputs.ST80_ET200SP_CM_4xIO_Link_3[25] := HwInputs.ST80_ET200SP_CM_4xIO_Link_3[25];
	PlcInputs.ST80_ET200SP_CM_4xIO_Link_3[26] := HwInputs.ST80_ET200SP_CM_4xIO_Link_3[26];
	PlcInputs.ST80_ET200SP_CM_4xIO_Link_3[27] := HwInputs.ST80_ET200SP_CM_4xIO_Link_3[27];
	PlcInputs.ST80_ET200SP_CM_4xIO_Link_3[28] := HwInputs.ST80_ET200SP_CM_4xIO_Link_3[28];
	PlcInputs.ST80_ET200SP_CM_4xIO_Link_3[29] := HwInputs.ST80_ET200SP_CM_4xIO_Link_3[29];
	PlcInputs.ST80_ET200SP_CM_4xIO_Link_3[30] := HwInputs.ST80_ET200SP_CM_4xIO_Link_3[30];
	PlcInputs.ST80_ET200SP_CM_4xIO_Link_3[31] := HwInputs.ST80_ET200SP_CM_4xIO_Link_3[31];
	PlcInputs.ST80_ET200SP_DI_16x24VDC_ST_1 := HwInputs.ST80_ET200SP_DI_16x24VDC_ST_1;
	PlcInputs.ST80_ET200SP_DI_16x24VDC_ST_2 := HwInputs.ST80_ET200SP_DI_16x24VDC_ST_2;
	PlcInputs.ST80_ET200SP_DI_16x24VDC_ST_3 := HwInputs.ST80_ET200SP_DI_16x24VDC_ST_3;
	PlcInputs.ST80_ET200SP_DI_16x24VDC_ST_4 := HwInputs.ST80_ET200SP_DI_16x24VDC_ST_4;
END_FUNCTION
